// Generated by scripts/make_plcsim_bench.py. Do not edit: rerun the script.
// Recorded force-travel curves from the Python model, the evaluation recipe of the study and the
// values the NumPy evaluation gives for the same samples. Read by FB_TestBench and FB_TestPlant.
//   X, F            samples of all curves, one after the other. A curve is CurveNPull pull samples
//                   followed by the same number of return samples, in the order they were taken.
//   Case..., Exp... replay cases 1..NCases: curve, evaluation mode, expected verdict, NOK code,
//                   elements (9 per case: FpG1 FrG1 FMean FHyst FpG2 FPeak XPeak FStep XStop) and
//                   envelope counts
//   Lim             16 limits per mode, index (mode - 1) * 16 + n, n in the order
//                   G1Lo G1Hi MeanLo MeanHi HystLo HystHi RetFMin G2Lo G2Hi PeakFLo PeakFHi PeakXMin PeakXMax StepLo StopXLo StopXHi
DATA_BLOCK "DB_TestData"
{ S7_Optimized_Access := 'TRUE' }
VERSION : 0.1
NON_RETAIN
   VAR
      NCurves : Int;
      NCases : Int;
      NSamples : Int;
      Tol : Real;   // N or mm, allowed difference of an element
      GoodCurve : Int;   // curve of the good unit in the station scenario
      BadCurve : Int;   // curve of the rejected unit in the station scenario
      GateX : Real;
      Gate2X : Real;
      PeakXLo : Real;
      PeakXHi : Real;
      StepSpan : Real;
      StopF : Real;
      EnvX0 : Real;
      EnvDx : Real;
      EnvN : Int;
      CurveStart : Array[0..15] of Int;
      CurveNPull : Array[0..15] of Int;
      CaseCurve : Array[1..32] of Int;
      CaseMode : Array[1..32] of Int;
      ExpOk : Array[1..32] of Bool;
      ExpNok : Array[1..32] of Int;
      ExpEnvViol : Array[1..32] of Int;
      ExpEnvNodes : Array[1..32] of Int;
      ExpFeat : Array[0..287] of Real;
      ExpFeatValid : Array[0..287] of Bool;
      Lim : Array[0..63] of Real;
      EnvLo : Array[0..63] of Real;
      EnvHi : Array[0..63] of Real;
      X : Array[0..5931] of Real;   // mm
      F : Array[0..5931] of Real;   // N
   END_VAR

BEGIN
   NCurves := 10;
   NCases := 14;
   NSamples := 5932;
   Tol := 0.001;
   GoodCurve := 0;
   BadCurve := 6;
   GateX := 3.0;
   Gate2X := 10.0;
   PeakXLo := 13.0;
   PeakXHi := 26.0;
   StepSpan := 2.0;
   StopF := 30.0;
   EnvX0 := 1.0;
   EnvDx := 0.5;
   EnvN := 55;
   CurveStart[0] := 0;
   CurveNPull[0] := 310;
   CurveStart[1] := 620;
   CurveNPull[1] := 313;
   CurveStart[2] := 1246;
   CurveNPull[2] := 250;
   CurveStart[3] := 1746;
   CurveNPull[3] := 310;
   CurveStart[4] := 2366;
   CurveNPull[4] := 311;
   CurveStart[5] := 2988;
   CurveNPull[5] := 309;
   CurveStart[6] := 3606;
   CurveNPull[6] := 311;
   CurveStart[7] := 4228;
   CurveNPull[7] := 250;
   CurveStart[8] := 4728;
   CurveNPull[8] := 291;
   CurveStart[9] := 5310;
   CurveNPull[9] := 311;
   CaseCurve[1] := 0;
   CaseMode[1] := 3;
   ExpOk[1] := TRUE;
   ExpNok[1] := 0;
   ExpEnvViol[1] := 0;
   ExpEnvNodes[1] := 55;
   ExpFeat[0] := 6.9821014;
   ExpFeatValid[0] := TRUE;
   ExpFeat[1] := 5.37568;
   ExpFeatValid[1] := TRUE;
   ExpFeat[2] := 6.1788907;
   ExpFeatValid[2] := TRUE;
   ExpFeat[3] := 1.6064217;
   ExpFeatValid[3] := TRUE;
   ExpFeat[4] := 10.845588;
   ExpFeatValid[4] := TRUE;
   ExpFeat[5] := 16.818577;
   ExpFeatValid[5] := TRUE;
   ExpFeat[6] := 19.848608;
   ExpFeatValid[6] := TRUE;
   ExpFeat[7] := 3.9388027;
   ExpFeatValid[7] := TRUE;
   ExpFeat[8] := 29.783041;
   ExpFeatValid[8] := TRUE;
   CaseCurve[2] := 1;
   CaseMode[2] := 3;
   ExpOk[2] := TRUE;
   ExpNok[2] := 0;
   ExpEnvViol[2] := 0;
   ExpEnvNodes[2] := 55;
   ExpFeat[9] := 7.205183;
   ExpFeatValid[9] := TRUE;
   ExpFeat[10] := 5.0210447;
   ExpFeatValid[10] := TRUE;
   ExpFeat[11] := 6.113114;
   ExpFeatValid[11] := TRUE;
   ExpFeat[12] := 2.1841383;
   ExpFeatValid[12] := TRUE;
   ExpFeat[13] := 11.2528515;
   ExpFeatValid[13] := TRUE;
   ExpFeat[14] := 17.15133;
   ExpFeatValid[14] := TRUE;
   ExpFeat[15] := 18.303595;
   ExpFeatValid[15] := TRUE;
   ExpFeat[16] := 4.152199;
   ExpFeatValid[16] := TRUE;
   ExpFeat[17] := 30.096466;
   ExpFeatValid[17] := TRUE;
   CaseCurve[3] := 2;
   CaseMode[3] := 3;
   ExpNok[3] := 2;
   ExpEnvViol[3] := 43;
   ExpEnvNodes[3] := 46;
   ExpFeat[18] := 4.183258;
   ExpFeatValid[18] := TRUE;
   ExpFeat[19] := 2.565676;
   ExpFeatValid[19] := TRUE;
   ExpFeat[20] := 3.374467;
   ExpFeatValid[20] := TRUE;
   ExpFeat[21] := 1.6175817;
   ExpFeatValid[21] := TRUE;
   ExpFeat[22] := 6.124597;
   ExpFeatValid[22] := TRUE;
   ExpFeat[23] := 40.227142;
   ExpFeatValid[23] := TRUE;
   ExpFeat[24] := 23.940363;
   ExpFeatValid[24] := TRUE;
   ExpFeat[25] := 0.0;
   ExpFeatValid[25] := TRUE;
   ExpFeat[26] := 23.785864;
   ExpFeatValid[26] := TRUE;
   CaseCurve[4] := 3;
   CaseMode[4] := 3;
   ExpNok[4] := 2;
   ExpEnvViol[4] := 0;
   ExpEnvNodes[4] := 55;
   ExpFeat[27] := 5.1918726;
   ExpFeatValid[27] := TRUE;
   ExpFeat[28] := 3.556863;
   ExpFeatValid[28] := TRUE;
   ExpFeat[29] := 4.3743677;
   ExpFeatValid[29] := TRUE;
   ExpFeat[30] := 1.6350094;
   ExpFeatValid[30] := TRUE;
   ExpFeat[31] := 9.031395;
   ExpFeatValid[31] := TRUE;
   ExpFeat[32] := 14.923322;
   ExpFeatValid[32] := TRUE;
   ExpFeat[33] := 19.814;
   ExpFeatValid[33] := TRUE;
   ExpFeat[34] := 3.9026327;
   ExpFeatValid[34] := TRUE;
   ExpFeat[35] := 29.81065;
   ExpFeatValid[35] := TRUE;
   CaseCurve[5] := 4;
   CaseMode[5] := 3;
   ExpNok[5] := 2;
   ExpEnvViol[5] := 17;
   ExpEnvNodes[5] := 55;
   ExpFeat[36] := 4.6947575;
   ExpFeatValid[36] := TRUE;
   ExpFeat[37] := 3.0623243;
   ExpFeatValid[37] := TRUE;
   ExpFeat[38] := 3.8785408;
   ExpFeatValid[38] := TRUE;
   ExpFeat[39] := 1.632433;
   ExpFeatValid[39] := TRUE;
   ExpFeat[40] := 8.425375;
   ExpFeatValid[40] := TRUE;
   ExpFeat[41] := 14.073351;
   ExpFeatValid[41] := TRUE;
   ExpFeat[42] := 19.786457;
   ExpFeatValid[42] := TRUE;
   ExpFeat[43] := 3.8736982;
   ExpFeatValid[43] := TRUE;
   ExpFeat[44] := 29.815647;
   ExpFeatValid[44] := TRUE;
   CaseCurve[6] := 5;
   CaseMode[6] := 3;
   ExpNok[6] := 3;
   ExpEnvViol[6] := 41;
   ExpEnvNodes[6] := 55;
   ExpFeat[45] := 10.499536;
   ExpFeatValid[45] := TRUE;
   ExpFeat[46] := 1.8700012;
   ExpFeatValid[46] := TRUE;
   ExpFeat[47] := 6.184768;
   ExpFeatValid[47] := TRUE;
   ExpFeat[48] := 8.629534;
   ExpFeatValid[48] := TRUE;
   ExpFeat[49] := 14.390507;
   ExpFeatValid[49] := TRUE;
   ExpFeat[50] := 20.330584;
   ExpFeatValid[50] := TRUE;
   ExpFeat[51] := 19.78603;
   ExpFeatValid[51] := TRUE;
   ExpFeat[52] := 3.8881645;
   ExpFeatValid[52] := TRUE;
   ExpFeat[53] := 29.722036;
   ExpFeatValid[53] := TRUE;
   CaseCurve[7] := 6;
   CaseMode[7] := 3;
   ExpNok[7] := 5;
   ExpEnvViol[7] := 41;
   ExpEnvNodes[7] := 55;
   ExpFeat[54] := 7.0127378;
   ExpFeatValid[54] := TRUE;
   ExpFeat[55] := 5.3387175;
   ExpFeatValid[55] := TRUE;
   ExpFeat[56] := 6.175728;
   ExpFeatValid[56] := TRUE;
   ExpFeat[57] := 1.67402;
   ExpFeatValid[57] := TRUE;
   ExpFeat[58] := 7.371472;
   ExpFeatValid[58] := TRUE;
   ExpFeat[59] := 8.326099;
   ExpFeatValid[59] := TRUE;
   ExpFeat[60] := 25.861488;
   ExpFeatValid[60] := TRUE;
   ExpFeat[61] := 0.032551765;
   ExpFeatValid[61] := TRUE;
   ExpFeat[62] := 29.877676;
   ExpFeatValid[62] := TRUE;
   CaseCurve[8] := 7;
   CaseMode[8] := 3;
   ExpNok[8] := 2;
   ExpEnvViol[8] := 43;
   ExpEnvNodes[8] := 46;
   ExpFeat[63] := 4.238579;
   ExpFeatValid[63] := TRUE;
   ExpFeat[64] := 2.6031868;
   ExpFeatValid[64] := TRUE;
   ExpFeat[65] := 3.420883;
   ExpFeatValid[65] := TRUE;
   ExpFeat[66] := 1.6353921;
   ExpFeatValid[66] := TRUE;
   ExpFeat[67] := 6.187137;
   ExpFeatValid[67] := TRUE;
   ExpFeat[68] := 41.858364;
   ExpFeatValid[68] := TRUE;
   ExpFeat[69] := 23.904263;
   ExpFeatValid[69] := TRUE;
   ExpFeat[70] := 0.0;
   ExpFeatValid[70] := TRUE;
   ExpFeat[71] := 23.727392;
   ExpFeatValid[71] := TRUE;
   CaseCurve[9] := 8;
   CaseMode[9] := 3;
   ExpNok[9] := 9;
   ExpEnvViol[9] := 1;
   ExpEnvNodes[9] := 55;
   ExpFeat[72] := 7.0128746;
   ExpFeatValid[72] := TRUE;
   ExpFeat[73] := 5.3684235;
   ExpFeatValid[73] := TRUE;
   ExpFeat[74] := 6.190649;
   ExpFeatValid[74] := TRUE;
   ExpFeat[75] := 1.6444514;
   ExpFeatValid[75] := TRUE;
   ExpFeat[76] := 10.856109;
   ExpFeatValid[76] := TRUE;
   ExpFeat[77] := 16.749855;
   ExpFeatValid[77] := TRUE;
   ExpFeat[78] := 19.791138;
   ExpFeatValid[78] := TRUE;
   ExpFeat[79] := 3.8845482;
   ExpFeatValid[79] := TRUE;
   ExpFeat[80] := 27.874788;
   ExpFeatValid[80] := TRUE;
   CaseCurve[10] := 9;
   CaseMode[10] := 3;
   ExpNok[10] := 2;
   ExpEnvViol[10] := 0;
   ExpEnvNodes[10] := 55;
   ExpFeat[81] := 6.2380857;
   ExpFeatValid[81] := TRUE;
   ExpFeat[82] := 2.573432;
   ExpFeatValid[82] := TRUE;
   ExpFeat[83] := 4.405759;
   ExpFeatValid[83] := TRUE;
   ExpFeat[84] := 3.6646535;
   ExpFeatValid[84] := TRUE;
   ExpFeat[85] := 10.107543;
   ExpFeatValid[85] := TRUE;
   ExpFeat[86] := 15.954138;
   ExpFeatValid[86] := TRUE;
   ExpFeat[87] := 19.8363;
   ExpFeatValid[87] := TRUE;
   ExpFeat[88] := 3.8773146;
   ExpFeatValid[88] := TRUE;
   ExpFeat[89] := 29.792097;
   ExpFeatValid[89] := TRUE;
   CaseCurve[11] := 9;
   CaseMode[11] := 2;
   ExpOk[11] := TRUE;
   ExpNok[11] := 0;
   ExpEnvViol[11] := 0;
   ExpEnvNodes[11] := 55;
   ExpFeat[90] := 6.2380857;
   ExpFeatValid[90] := TRUE;
   ExpFeat[91] := 2.573432;
   ExpFeatValid[91] := TRUE;
   ExpFeat[92] := 4.405759;
   ExpFeatValid[92] := TRUE;
   ExpFeat[93] := 3.6646535;
   ExpFeatValid[93] := TRUE;
   ExpFeat[94] := 10.107543;
   ExpFeatValid[94] := TRUE;
   ExpFeat[95] := 15.954138;
   ExpFeatValid[95] := TRUE;
   ExpFeat[96] := 19.8363;
   ExpFeatValid[96] := TRUE;
   ExpFeat[97] := 3.8773146;
   ExpFeatValid[97] := TRUE;
   ExpFeat[98] := 29.792097;
   ExpFeatValid[98] := TRUE;
   CaseCurve[12] := 8;
   CaseMode[12] := 1;
   ExpOk[12] := TRUE;
   ExpNok[12] := 0;
   ExpEnvViol[12] := 1;
   ExpEnvNodes[12] := 55;
   ExpFeat[99] := 7.0128746;
   ExpFeatValid[99] := TRUE;
   ExpFeat[100] := 5.3684235;
   ExpFeatValid[100] := TRUE;
   ExpFeat[101] := 6.190649;
   ExpFeatValid[101] := TRUE;
   ExpFeat[102] := 1.6444514;
   ExpFeatValid[102] := TRUE;
   ExpFeat[103] := 10.856109;
   ExpFeatValid[103] := TRUE;
   ExpFeat[104] := 16.749855;
   ExpFeatValid[104] := TRUE;
   ExpFeat[105] := 19.791138;
   ExpFeatValid[105] := TRUE;
   ExpFeat[106] := 3.8845482;
   ExpFeatValid[106] := TRUE;
   ExpFeat[107] := 27.874788;
   ExpFeatValid[107] := TRUE;
   CaseCurve[13] := 0;
   CaseMode[13] := 4;
   ExpOk[13] := TRUE;
   ExpNok[13] := 0;
   ExpEnvViol[13] := 0;
   ExpEnvNodes[13] := 55;
   ExpFeat[108] := 6.9821014;
   ExpFeatValid[108] := TRUE;
   ExpFeat[109] := 5.37568;
   ExpFeatValid[109] := TRUE;
   ExpFeat[110] := 6.1788907;
   ExpFeatValid[110] := TRUE;
   ExpFeat[111] := 1.6064217;
   ExpFeatValid[111] := TRUE;
   ExpFeat[112] := 10.845588;
   ExpFeatValid[112] := TRUE;
   ExpFeat[113] := 16.818577;
   ExpFeatValid[113] := TRUE;
   ExpFeat[114] := 19.848608;
   ExpFeatValid[114] := TRUE;
   ExpFeat[115] := 3.9388027;
   ExpFeatValid[115] := TRUE;
   ExpFeat[116] := 29.783041;
   ExpFeatValid[116] := TRUE;
   CaseCurve[14] := 3;
   CaseMode[14] := 4;
   ExpOk[14] := TRUE;
   ExpNok[14] := 0;
   ExpEnvViol[14] := 0;
   ExpEnvNodes[14] := 55;
   ExpFeat[117] := 5.1918726;
   ExpFeatValid[117] := TRUE;
   ExpFeat[118] := 3.556863;
   ExpFeatValid[118] := TRUE;
   ExpFeat[119] := 4.3743677;
   ExpFeatValid[119] := TRUE;
   ExpFeat[120] := 1.6350094;
   ExpFeatValid[120] := TRUE;
   ExpFeat[121] := 9.031395;
   ExpFeatValid[121] := TRUE;
   ExpFeat[122] := 14.923322;
   ExpFeatValid[122] := TRUE;
   ExpFeat[123] := 19.814;
   ExpFeatValid[123] := TRUE;
   ExpFeat[124] := 3.9026327;
   ExpFeatValid[124] := TRUE;
   ExpFeat[125] := 29.81065;
   ExpFeatValid[125] := TRUE;
   Lim[9] := 15.241609;
   Lim[10] := 18.417305;
   Lim[16] := 5.896105;
   Lim[17] := 8.38203;
   Lim[23] := 9.4181;
   Lim[24] := 12.402887;
   Lim[25] := 14.982571;
   Lim[26] := 18.676344;
   Lim[27] := 17.139359;
   Lim[28] := 22.516165;
   Lim[29] := 2.9451215;
   Lim[30] := 28.690018;
   Lim[31] := 30.871372;
   Lim[34] := 5.186474;
   Lim[35] := 7.2080727;
   Lim[36] := -0.5455249;
   Lim[37] := 3.975223;
   Lim[38] := 1.0;
   Lim[39] := 9.212741;
   Lim[40] := 12.608247;
   Lim[41] := 14.728432;
   Lim[42] := 18.930483;
   Lim[43] := 16.769424;
   Lim[44] := 22.886099;
   Lim[45] := 2.8110514;
   Lim[46] := 28.539938;
   Lim[47] := 31.021452;
   EnvLo[0] := 4.5024867;
   EnvHi[0] := 9.917023;
   EnvLo[1] := 4.5624857;
   EnvHi[1] := 9.98225;
   EnvLo[2] := 4.530773;
   EnvHi[2] := 9.992803;
   EnvLo[3] := 4.5635424;
   EnvHi[3] := 10.004515;
   EnvLo[4] := 4.573186;
   EnvHi[4] := 10.029344;
   EnvLo[5] := 4.617667;
   EnvHi[5] := 10.026862;
   EnvLo[6] := 4.6239376;
   EnvHi[6] := 10.070514;
   EnvLo[7] := 4.670679;
   EnvHi[7] := 10.102605;
   EnvLo[8] := 4.725596;
   EnvHi[8] := 12.041139;
   EnvLo[9] := 4.700003;
   EnvHi[9] := 12.557893;
   EnvLo[10] := 4.8820324;
   EnvHi[10] := 12.779339;
   EnvLo[11] := 4.926072;
   EnvHi[11] := 12.91771;
   EnvLo[12] := 5.163019;
   EnvHi[12] := 13.360822;
   EnvLo[13] := 5.6595745;
   EnvHi[13] := 13.471234;
   EnvLo[14] := 7.878658;
   EnvHi[14] := 13.533369;
   EnvLo[15] := 8.020163;
   EnvHi[15] := 13.642666;
   EnvLo[16] := 8.08159;
   EnvHi[16] := 13.729599;
   EnvLo[17] := 8.207902;
   EnvHi[17] := 13.860825;
   EnvLo[18] := 8.30263;
   EnvHi[18] := 13.911284;
   EnvLo[19] := 8.350869;
   EnvHi[19] := 13.990431;
   EnvLo[20] := 8.425625;
   EnvHi[20] := 14.0966015;
   EnvLo[21] := 8.550419;
   EnvHi[21] := 14.182879;
   EnvLo[22] := 8.607436;
   EnvHi[22] := 14.296827;
   EnvLo[23] := 8.764787;
   EnvHi[23] := 14.390328;
   EnvLo[24] := 8.845735;
   EnvHi[24] := 14.4539795;
   EnvLo[25] := 8.9147835;
   EnvHi[25] := 14.551714;
   EnvLo[26] := 8.99205;
   EnvHi[26] := 14.698472;
   EnvLo[27] := 9.068602;
   EnvHi[27] := 15.185006;
   EnvLo[28] := 9.331687;
   EnvHi[28] := 15.688478;
   EnvLo[29] := 9.416069;
   EnvHi[29] := 16.23098;
   EnvLo[30] := 9.513143;
   EnvHi[30] := 16.795422;
   EnvLo[31] := 9.665618;
   EnvHi[31] := 17.309069;
   EnvLo[32] := 10.123489;
   EnvHi[32] := 17.854668;
   EnvLo[33] := 10.642103;
   EnvHi[33] := 18.362646;
   EnvLo[34] := 11.14989;
   EnvHi[34] := 18.931261;
   EnvLo[35] := 11.027167;
   EnvHi[35] := 18.921373;
   EnvLo[36] := 10.830289;
   EnvHi[36] := 19.396362;
   EnvLo[37] := 10.428676;
   EnvHi[37] := 19.986576;
   EnvLo[38] := 10.27112;
   EnvHi[38] := 19.496552;
   EnvLo[39] := 10.313659;
   EnvHi[39] := 19.897247;
   EnvLo[40] := 10.363278;
   EnvHi[40] := 19.346785;
   EnvLo[41] := 10.468162;
   EnvHi[41] := 18.766773;
   EnvLo[42] := 10.585302;
   EnvHi[42] := 16.553541;
   EnvLo[43] := 10.677869;
   EnvHi[43] := 16.354622;
   EnvLo[44] := 10.748317;
   EnvHi[44] := 16.457827;
   EnvLo[45] := 10.8695135;
   EnvHi[45] := 16.512941;
   EnvLo[46] := 10.998811;
   EnvHi[46] := 16.617954;
   EnvLo[47] := 11.099038;
   EnvHi[47] := 16.769545;
   EnvLo[48] := 11.214338;
   EnvHi[48] := 16.847044;
   EnvLo[49] := 11.278554;
   EnvHi[49] := 16.997396;
   EnvLo[50] := 11.41541;
   EnvHi[50] := 17.054838;
   EnvLo[51] := 11.506263;
   EnvHi[51] := 17.213253;
   EnvLo[52] := 11.623229;
   EnvHi[52] := 17.348417;
   EnvLo[53] := 11.713954;
   EnvHi[53] := 17.397055;
   EnvLo[54] := 11.844806;
   EnvHi[54] := 17.536877;
   X[1] := -0.0033742767;
   X[2] := 0.10472685;
   X[3] := 0.19745024;
   X[4] := 0.29981726;
   X[5] := 0.39700347;
   X[6] := 0.49491304;
   X[7] := 0.6008226;
   X[8] := 0.6972801;
   X[9] := 0.7991843;
   X[10] := 0.90281725;
   X[11] := 0.99573755;
   X[12] := 1.0995567;
   X[13] := 1.1978173;
   X[14] := 1.2951844;
   X[15] := 1.3980939;
   X[16] := 1.4998226;
   X[17] := 1.5985514;
   X[18] := 1.7018226;
   X[19] := 1.8003706;
   X[20] := 1.8912854;
   X[21] := 1.999562;
   X[22] := 2.0993705;
   X[23] := 2.1909237;
   X[24] := 2.2984662;
   X[25] := 2.3891046;
   X[26] := 2.4932854;
   X[27] := 2.601009;
   X[28] := 2.6959238;
   X[29] := 2.796014;
   X[30] := 2.894743;
   X[31] := 2.9955568;
   X[32] := 3.092743;
   X[33] := 3.1978333;
   X[34] := 3.292743;
   X[35] := 3.3987377;
   X[36] := 3.4987428;
   X[37] := 3.59511;
   X[38] := 3.6955674;
   X[39] := 3.7989292;
   X[40] := 3.8956633;
   X[41] := 3.9927535;
   X[42] := 4.0977483;
   X[43] := 4.197296;
   X[44] := 4.292573;
   X[45] := 4.399477;
   X[46] := 4.4931207;
   X[47] := 4.593658;
   X[48] := 4.6908493;
   X[49] := 4.7944875;
   X[50] := 4.8961205;
   X[51] := 4.9969397;
   X[52] := 5.094764;
   X[53] := 5.18994;
   X[54] := 5.2910357;
   X[55] := 5.394844;
   X[56] := 5.489573;
   X[57] := 5.5893974;
   X[58] := 5.6894984;
   X[59] := 5.7891207;
   X[60] := 5.893126;
   X[61] := 5.989312;
   X[62] := 6.076935;
   X[63] := 6.1627493;
   X[64] := 6.2443776;
   X[65] := 6.328378;
   X[66] := 6.4094586;
   X[67] := 6.5168147;
   X[68] := 6.6171765;
   X[69] := 6.718815;
   X[70] := 6.8094583;
   X[71] := 6.9220915;
   X[72] := 7.0171022;
   X[73] := 7.1126394;
   X[74] := 7.213565;
   X[75] := 7.3112035;
   X[76] := 7.4117403;
   X[77] := 7.511751;
   X[78] := 7.606661;
   X[79] := 7.708384;
   X[80] := 7.81248;
   X[81] := 7.9090276;
   X[82] := 8.005486;
   X[83] := 8.110033;
   X[84] := 8.2134;
   X[85] := 8.307496;
   X[86] := 8.410586;
   X[87] := 8.505591;
   X[88] := 8.600773;
   X[89] := 8.702959;
   X[90] := 8.809416;
   X[91] := 8.908698;
   X[92] := 8.999699;
   X[93] := 9.103602;
   X[94] := 9.201704;
   X[95] := 9.301433;
   X[96] := 9.39789;
   X[97] := 9.503613;
   X[98] := 9.601155;
   X[99] := 9.699528;
   X[100] := 9.802805;
   X[101] := 9.89989;
   X[102] := 10.003895;
   X[103] := 10.098449;
   X[104] := 10.201262;
   X[105] := 10.298172;
   X[106] := 10.399454;
   X[107] := 10.497454;
   X[108] := 10.592826;
   X[109] := 10.699917;
   X[110] := 10.798554;
   X[111] := 10.89847;
   X[112] := 10.996193;
   X[113] := 11.098837;
   X[114] := 11.192114;
   X[115] := 11.287757;
   X[116] := 11.391119;
   X[117] := 11.496119;
   X[118] := 11.592933;
   X[119] := 11.693028;
   X[120] := 11.786496;
   X[121] := 11.891943;
   X[122] := 11.991592;
   X[123] := 12.0868635;
   X[124] := 12.186582;
   X[125] := 12.291321;
   X[126] := 12.380411;
   X[127] := 12.48514;
   X[128] := 12.584327;
   X[129] := 12.683965;
   X[130] := 12.787603;
   X[131] := 12.888337;
   X[132] := 12.989885;
   X[133] := 13.08306;
   X[134] := 13.187704;
   X[135] := 13.284523;
   X[136] := 13.3848;
   X[137] := 13.487896;
   X[138] := 13.587353;
   X[139] := 13.678811;
   X[140] := 13.784454;
   X[141] := 13.882715;
   X[142] := 13.981008;
   X[143] := 14.078545;
   X[144] := 14.183087;
   X[145] := 14.28164;
   X[146] := 14.38038;
   X[147] := 14.475013;
   X[148] := 14.574927;
   X[149] := 14.682922;
   X[150] := 14.780104;
   X[151] := 14.878199;
   X[152] := 14.975023;
   X[153] := 15.076039;
   X[154] := 15.17287;
   X[155] := 15.271434;
   X[156] := 15.363907;
   X[157] := 15.460098;
   X[158] := 15.557104;
   X[159] := 15.660487;
   X[160] := 15.751045;
   X[161] := 15.851062;
   X[162] := 15.951705;
   X[163] := 16.053541;
   X[164] := 16.149647;
   X[165] := 16.244019;
   X[166] := 16.34385;
   X[167] := 16.440685;
   X[168] := 16.537062;
   X[169] := 16.62862;
   X[170] := 16.734083;
   X[171] := 16.83637;
   X[172] := 16.92229;
   X[173] := 17.019585;
   X[174] := 17.119505;
   X[175] := 17.217972;
   X[176] := 17.316803;
   X[177] := 17.418;
   X[178] := 17.508282;
   X[179] := 17.611292;
   X[180] := 17.70858;
   X[181] := 17.800692;
   X[182] := 17.902872;
   X[183] := 17.99408;
   X[184] := 18.09909;
   X[185] := 18.191565;
   X[186] := 18.287483;
   X[187] := 18.387772;
   X[188] := 18.49033;
   X[189] := 18.585798;
   X[190] := 18.676447;
   X[191] := 18.777182;
   X[192] := 18.874111;
   X[193] := 18.979118;
   X[194] := 19.070032;
   X[195] := 19.165964;
   X[196] := 19.270985;
   X[197] := 19.360996;
   X[198] := 19.462011;
   X[199] := 19.55457;
   X[200] := 19.65848;
   X[201] := 19.755777;
   X[202] := 19.848608;
   X[203] := 19.970793;
   X[204] := 20.087416;
   X[205] := 20.211292;
   X[206] := 20.32783;
   X[207] := 20.445093;
   X[208] := 20.557806;
   X[209] := 20.648077;
   X[210] := 20.741636;
   X[211] := 20.84809;
   X[212] := 20.953089;
   X[213] := 21.043913;
   X[214] := 21.147093;
   X[215] := 21.24119;
   X[216] := 21.348913;
   X[217] := 21.449648;
   X[218] := 21.545195;
   X[219] := 21.634748;
   X[220] := 21.745749;
   X[221] := 21.841301;
   X[222] := 21.946121;
   X[223] := 22.040205;
   X[224] := 22.143402;
   X[225] := 22.240217;
   X[226] := 22.341042;
   X[227] := 22.44068;
   X[228] := 22.53859;
   X[229] := 22.634499;
   X[230] := 22.738136;
   X[231] := 22.838509;
   X[232] := 22.941322;
   X[233] := 23.042967;
   X[234] := 23.129976;
   X[235] := 23.239418;
   X[236] := 23.335434;
   X[237] := 23.430067;
   X[238] := 23.531801;
   X[239] := 23.641802;
   X[240] := 23.734535;
   X[241] := 23.835356;
   X[242] := 23.933903;
   X[243] := 24.02927;
   X[244] := 24.133179;
   X[245] := 24.232546;
   X[246] := 24.332918;
   X[247] := 24.43128;
   X[248] := 24.52801;
   X[249] := 24.624918;
   X[250] := 24.728653;
   X[251] := 24.823557;
   X[252] := 24.925116;
   X[253] := 25.026297;
   X[254] := 25.123116;
   X[255] := 25.230398;
   X[256] := 25.325674;
   X[257] := 25.426765;
   X[258] := 25.523584;
   X[259] := 25.621408;
   X[260] := 25.71895;
   X[261] := 25.820227;
   X[262] := 25.919882;
   X[263] := 26.019594;
   X[264] := 26.116701;
   X[265] := 26.216702;
   X[266] := 26.315063;
   X[267] := 26.42161;
   X[268] := 26.524881;
   X[269] := 26.622345;
   X[270] := 26.714718;
   X[271] := 26.815802;
   X[272] := 26.917803;
   X[273] := 27.014627;
   X[274] := 27.115812;
   X[275] := 27.214813;
   X[276] := 27.312366;
   X[277] := 27.413908;
   X[278] := 27.51119;
   X[279] := 27.612286;
   X[280] := 27.709558;
   X[281] := 27.811739;
   X[282] := 27.911112;
   X[283] := 28.007027;
   X[284] := 28.111387;
   X[285] := 28.199669;
   X[286] := 28.301207;
   X[287] := 28.40676;
   X[288] := 28.508398;
   X[289] := 28.60403;
   X[290] := 28.701595;
   X[291] := 28.8095;
   X[292] := 28.900776;
   X[293] := 29.00051;
   X[294] := 29.101877;
   X[295] := 29.200064;
   X[296] := 29.301426;
   X[297] := 29.398798;
   X[298] := 29.500973;
   X[299] := 29.572319;
   X[300] := 29.6092;
   X[301] := 29.646812;
   X[302] := 29.686869;
   X[303] := 29.716297;
   X[304] := 29.758177;
   X[305] := 29.799242;
   X[306] := 29.837845;
   X[307] := 29.867996;
   X[308] := 29.91243;
   X[309] := 29.94758;
   X[310] := 29.943314;
   X[311] := 29.928886;
   X[312] := 29.886644;
   X[313] := 29.850302;
   X[314] := 29.813248;
   X[315] := 29.77291;
   X[316] := 29.739481;
   X[317] := 29.693878;
   X[318] := 29.666807;
   X[319] := 29.625662;
   X[320] := 29.588596;
   X[321] := 29.545658;
   X[322] := 29.446291;
   X[323] := 29.346828;
   X[324] := 29.248291;
   X[325] := 29.144827;
   X[326] := 29.049004;
   X[327] := 28.937727;
   X[328] := 28.847637;
   X[329] := 28.75453;
   X[330] := 28.642721;
   X[331] := 28.549807;
   X[332] := 28.448168;
   X[333] := 28.348167;
   X[334] := 28.251705;
   X[335] := 28.151072;
   X[336] := 28.05543;
   X[337] := 27.9487;
   X[338] := 27.857418;
   X[339] := 27.751062;
   X[340] := 27.654417;
   X[341] := 27.556412;
   X[342] := 27.45969;
   X[343] := 27.360954;
   X[344] := 27.257498;
   X[345] := 27.15513;
   X[346] := 27.059216;
   X[347] := 26.958311;
   X[348] := 26.85785;
   X[349] := 26.761482;
   X[350] := 26.654758;
   X[351] := 26.5573;
   X[352] := 26.460743;
   X[353] := 26.360561;
   X[354] := 26.257103;
   X[355] := 26.160013;
   X[356] := 26.06664;
   X[357] := 25.96328;
   X[358] := 25.863731;
   X[359] := 25.76454;
   X[360] := 25.668083;
   X[361] := 25.56563;
   X[362] := 25.464897;
   X[363] := 25.367987;
   X[364] := 25.26344;
   X[365] := 25.167982;
   X[366] := 25.070257;
   X[367] := 24.966524;
   X[368] := 24.871796;
   X[369] := 24.767876;
   X[370] := 24.67279;
   X[371] := 24.576056;
   X[372] := 24.471146;
   X[373] := 24.368502;
   X[374] := 24.26669;
   X[375] := 24.170046;
   X[376] := 24.073677;
   X[377] := 23.97786;
   X[378] := 23.87113;
   X[379] := 23.777668;
   X[380] := 23.676853;
   X[381] := 23.576395;
   X[382] := 23.480204;
   X[383] := 23.375023;
   X[384] := 23.272934;
   X[385] := 23.17702;
   X[386] := 23.081102;
   X[387] := 22.978556;
   X[388] := 22.88028;
   X[389] := 22.779646;
   X[390] := 22.677635;
   X[391] := 22.582449;
   X[392] := 22.482183;
   X[393] := 22.376087;
   X[394] := 22.28681;
   X[395] := 22.185173;
   X[396] := 22.084444;
   X[397] := 21.981167;
   X[398] := 21.891161;
   X[399] := 21.780619;
   X[400] := 21.684343;
   X[401] := 21.589523;
   X[402] := 21.48388;
   X[403] := 21.391508;
   X[404] := 21.285975;
   X[405] := 21.187326;
   X[406] := 21.08787;
   X[407] := 20.986044;
   X[408] := 20.88931;
   X[409] := 20.790411;
   X[410] := 20.692492;
   X[411] := 20.591034;
   X[412] := 20.4904;
   X[413] := 20.394842;
   X[414] := 20.293018;
   X[415] := 20.197294;
   X[416] := 20.102022;
   X[417] := 19.994108;
   X[418] := 19.893831;
   X[419] := 19.797018;
   X[420] := 19.694916;
   X[421] := 19.590475;
   X[422] := 19.501102;
   X[423] := 19.397188;
   X[424] := 19.298725;
   X[425] := 19.19691;
   X[426] := 19.100178;
   X[427] := 18.99881;
   X[428] := 18.902714;
   X[429] := 18.797997;
   X[430] := 18.700708;
   X[431] := 18.604261;
   X[432] := 18.502884;
   X[433] := 18.39889;
   X[434] := 18.303162;
   X[435] := 18.206156;
   X[436] := 18.103241;
   X[437] := 17.99897;
   X[438] := 17.907688;
   X[439] := 17.802235;
   X[440] := 17.704773;
   X[441] := 17.608416;
   X[442] := 17.508411;
   X[443] := 17.407219;
   X[444] := 17.30849;
   X[445] := 17.209394;
   X[446] := 17.109943;
   X[447] := 17.011847;
   X[448] := 16.906948;
   X[449] := 16.809395;
   X[450] := 16.708118;
   X[451] := 16.613565;
   X[452] := 16.507107;
   X[453] := 16.412107;
   X[454] := 16.31701;
   X[455] := 16.208832;
   X[456] := 16.112278;
   X[457] := 16.011374;
   X[458] := 15.918001;
   X[459] := 15.814639;
   X[460] := 15.7179;
   X[461] := 15.617182;
   X[462] := 15.515448;
   X[463] := 15.413996;
   X[464] := 15.3189;
   X[465] := 15.21989;
   X[466] := 15.117075;
   X[467] := 15.018708;
   X[468] := 14.91516;
   X[469] := 14.81798;
   X[470] := 14.721788;
   X[471] := 14.619889;
   X[472] := 14.519878;
   X[473] := 14.4160595;
   X[474] := 14.324873;
   X[475] := 14.220602;
   X[476] := 14.128693;
   X[477] := 14.019857;
   X[478] := 13.914687;
   X[479] := 13.827314;
   X[480] := 13.7215;
   X[481] := 13.626677;
   X[482] := 13.521501;
   X[483] := 13.424581;
   X[484] := 13.327847;
   X[485] := 13.228756;
   X[486] := 13.133394;
   X[487] := 13.029112;
   X[488] := 12.930293;
   X[489] := 12.828841;
   X[490] := 12.727287;
   X[491] := 12.62883;
   X[492] := 12.531464;
   X[493] := 12.429921;
   X[494] := 12.327181;
   X[495] := 12.229639;
   X[496] := 12.131453;
   X[497] := 12.032723;
   X[498] := 11.925458;
   X[499] := 11.833815;
   X[500] := 11.732442;
   X[501] := 11.633894;
   X[502] := 11.536803;
   X[503] := 11.433075;
   X[504] := 11.328346;
   X[505] := 11.23716;
   X[506] := 11.135245;
   X[507] := 11.032245;
   X[508] := 10.939425;
   X[509] := 10.837878;
   X[510] := 10.737963;
   X[511] := 10.632873;
   X[512] := 10.537234;
   X[513] := 10.437139;
   X[514] := 10.339868;
   X[515] := 10.24041;
   X[516] := 10.143681;
   X[517] := 10.045037;
   X[518] := 9.939037;
   X[519] := 9.833128;
   X[520] := 9.744676;
   X[521] := 9.642303;
   X[522] := 9.540303;
   X[523] := 9.441941;
   X[524] := 9.343032;
   X[525] := 9.2415695;
   X[526] := 9.141931;
   X[527] := 9.047192;
   X[528] := 8.943649;
   X[529] := 8.843558;
   X[530] := 8.747462;
   X[531] := 8.645282;
   X[532] := 8.554914;
   X[533] := 8.446638;
   X[534] := 8.344186;
   X[535] := 8.247452;
   X[536] := 8.145633;
   X[537] := 8.051356;
   X[538] := 7.9505424;
   X[539] := 7.854803;
   X[540] := 7.749255;
   X[541] := 7.6534357;
   X[542] := 7.5542603;
   X[543] := 7.453893;
   X[544] := 7.3493347;
   X[545] := 7.2504253;
   X[546] := 7.1519732;
   X[547] := 7.054606;
   X[548] := 6.9581485;
   X[549] := 6.8538775;
   X[550] := 6.7531433;
   X[551] := 6.657409;
   X[552] := 6.5563293;
   X[553] := 6.4607816;
   X[554] := 6.3632812;
   X[555] := 6.274286;
   X[556] := 6.1935673;
   X[557] := 6.108753;
   X[558] := 6.03021;
   X[559] := 5.9339066;
   X[560] := 5.8310876;
   X[561] := 5.731545;
   X[562] := 5.6369066;
   X[563] := 5.531364;
   X[564] := 5.437353;
   X[565] := 5.337811;
   X[566] := 5.2275395;
   X[567] := 5.126901;
   X[568] := 5.03872;
   X[569] := 4.9384384;
   X[570] := 4.8375287;
   X[571] := 4.739082;
   X[572] := 4.634901;
   X[573] := 4.5331616;
   X[574] := 4.4404383;
   X[575] := 4.329167;
   X[576] := 4.233348;
   X[577] := 4.1344438;
   X[578] := 4.0365286;
   X[579] := 3.9392576;
   X[580] := 3.834167;
   X[581] := 3.7369862;
   X[582] := 3.633433;
   X[583] := 3.5345287;
   X[584] := 3.4394383;
   X[585] := 3.3372576;
   X[586] := 3.2332575;
   X[587] := 3.140433;
   X[588] := 3.043066;
   X[589] := 2.9320712;
   X[590] := 2.8413372;
   X[591] := 2.7396085;
   X[592] := 2.6366086;
   X[593] := 2.5347893;
   X[594] := 2.441518;
   X[595] := 2.342518;
   X[596] := 2.2378001;
   X[597] := 2.1382415;
   X[598] := 2.034066;
   X[599] := 1.9376031;
   X[600] := 1.8358798;
   X[601] := 1.7395127;
   X[602] := 1.6385127;
   X[603] := 1.540151;
   X[604] := 1.4401511;
   X[605] := 1.3368851;
   X[606] := 1.2400553;
   X[607] := 1.133151;
   X[608] := 1.0449648;
   X[609] := 0.939784;
   X[610] := 0.8416882;
   X[611] := 0.7337893;
   X[612] := 0.6410499;
   X[613] := 0.5402415;
   X[614] := 0.43896484;
   X[615] := 0.34032118;
   X[616] := 0.23696484;
   X[617] := 0.14223076;
   X[618] := 0.03723076;
   X[619] := 0.07943374;
   X[621] := 0.058969617;
   X[622] := 0.1601451;
   X[623] := 0.25842172;
   X[624] := 0.36087385;
   X[625] := 0.45877805;
   X[626] := 0.5548792;
   X[627] := 0.6574271;
   X[628] := 0.75815046;
   X[629] := 0.85487384;
   X[630] := 0.9517888;
   X[631] := 1.053975;
   X[632] := 1.1582409;
   X[633] := 1.2541559;
   X[634] := 1.3572463;
   X[635] := 1.4556025;
   X[636] := 1.5523367;
   X[637] := 1.6556187;
   X[638] := 1.7556983;
   X[639] := 1.8526186;
   X[640] := 1.9547037;
   X[641] := 2.0571558;
   X[642] := 2.1517036;
   X[643] := 2.2567995;
   X[644] := 2.3577092;
   X[645] := 2.4552517;
   X[646] := 2.5556185;
   X[647] := 2.6554377;
   X[648] := 2.7547994;
   X[649] := 2.850161;
   X[650] := 2.9497144;
   X[651] := 3.0517995;
   X[652] := 3.1496186;
   X[653] := 3.257076;
   X[654] := 3.3558953;
   X[655] := 3.4521666;
   X[656] := 3.5518048;
   X[657] := 3.653624;
   X[658] := 3.7534378;
   X[659] := 3.852991;
   X[660] := 3.9552622;
   X[661] := 4.04972;
   X[662] := 4.1526294;
   X[663] := 4.255996;
   X[664] := 4.3528047;
   X[665] := 4.4510016;
   X[666] := 4.5480866;
   X[667] := 4.6492677;
   X[668] := 4.7482677;
   X[669] := 4.853805;
   X[670] := 4.9477253;
   X[671] := 5.051906;
   X[672] := 5.151358;
   X[673] := 5.2348957;
   X[674] := 5.3198113;
   X[675] := 5.4007053;
   X[676] := 5.4895253;
   X[677] := 5.573419;
   X[678] := 5.673228;
   X[679] := 5.771866;
   X[680] := 5.871143;
   X[681] := 5.969329;
   X[682] := 6.072978;
   X[683] := 6.165616;
   X[684] := 6.2763395;
   X[685] := 6.37834;
   X[686] := 6.4693394;
   X[687] := 6.5714407;
   X[688] := 6.6652493;
   X[689] := 6.770627;
   X[690] := 6.8630843;
   X[691] := 6.9633555;
   X[692] := 7.0697227;
   X[693] := 7.168909;
   X[694] := 7.2685523;
   X[695] := 7.3637385;
   X[696] := 7.4669037;
   X[697] := 7.563648;
   X[698] := 7.6645527;
   X[699] := 7.7610154;
   X[700] := 7.8674674;
   X[701] := 7.9631057;
   X[702] := 8.063478;
   X[703] := 8.159749;
   X[704] := 8.254574;
   X[705] := 8.355664;
   X[706] := 8.462856;
   X[707] := 8.553574;
   X[708] := 8.662393;
   X[709] := 8.762766;
   X[710] := 8.8588505;
   X[711] := 8.952951;
   X[712] := 9.056047;
   X[713] := 9.15259;
   X[714] := 9.251148;
   X[715] := 9.357691;
   X[716] := 9.453968;
   X[717] := 9.555329;
   X[718] := 9.654702;
   X[719] := 9.75134;
   X[720] := 9.855978;
   X[721] := 9.954888;
   X[722] := 10.04817;
   X[723] := 10.15099;
   X[724] := 10.252255;
   X[725] := 10.3547125;
   X[726] := 10.451904;
   X[727] := 10.551271;
   X[728] := 10.646809;
   X[729] := 10.748909;
   X[730] := 10.853186;
   X[731] := 10.952457;
   X[732] := 11.050553;
   X[733] := 11.14801;
   X[734] := 11.246378;
   X[735] := 11.350468;
   X[736] := 11.444835;
   X[737] := 11.546383;
   X[738] := 11.644745;
   X[739] := 11.748659;
   X[740] := 11.844665;
   X[741] := 11.942393;
   X[742] := 12.038213;
   X[743] := 12.13958;
   X[744] := 12.245122;
   X[745] := 12.339048;
   X[746] := 12.439409;
   X[747] := 12.540957;
   X[748] := 12.639862;
   X[749] := 12.740053;
   X[750] := 12.837516;
   X[751] := 12.932607;
   X[752] := 13.040059;
   X[753] := 13.139059;
   X[754] := 13.238154;
   X[755] := 13.338431;
   X[756] := 13.4359;
   X[757] := 13.5304575;
   X[758] := 13.635559;
   X[759] := 13.72675;
   X[760] := 13.818857;
   X[761] := 13.918681;
   X[762] := 14.016246;
   X[763] := 14.117352;
   X[764] := 14.217459;
   X[765] := 14.311023;
   X[766] := 14.407762;
   X[767] := 14.50431;
   X[768] := 14.610332;
   X[769] := 14.701975;
   X[770] := 14.796544;
   X[771] := 14.899007;
   X[772] := 14.994475;
   X[773] := 15.085858;
   X[774] := 15.194316;
   X[775] := 15.28988;
   X[776] := 15.3827095;
   X[777] := 15.478273;
   X[778] := 15.579289;
   X[779] := 15.676763;
   X[780] := 15.776773;
   X[781] := 15.875156;
   X[782] := 15.973704;
   X[783] := 16.068811;
   X[784] := 16.163736;
   X[785] := 16.2553;
   X[786] := 16.359764;
   X[787] := 16.457323;
   X[788] := 16.552242;
   X[789] := 16.653168;
   X[790] := 16.743004;
   X[791] := 16.841015;
   X[792] := 16.939758;
   X[793] := 17.037136;
   X[794] := 17.140327;
   X[795] := 17.235802;
   X[796] := 17.331541;
   X[797] := 17.428104;
   X[798] := 17.52593;
   X[799] := 17.631126;
   X[800] := 17.718876;
   X[801] := 17.81943;
   X[802] := 17.915802;
   X[803] := 18.00819;
   X[804] := 18.111834;
   X[805] := 18.202488;
   X[806] := 18.303595;
   X[807] := 18.407286;
   X[808] := 18.52944;
   X[809] := 18.65905;
   X[810] := 18.7763;
   X[811] := 18.901001;
   X[812] := 19.0094;
   X[813] := 19.106045;
   X[814] := 19.20614;
   X[815] := 19.303415;
   X[816] := 19.40779;
   X[817] := 19.507235;
   X[818] := 19.609697;
   X[819] := 19.70224;
   X[820] := 19.802341;
   X[821] := 19.900156;
   X[822] := 20.002895;
   X[823] := 20.102533;
   X[824] := 20.202618;
   X[825] := 20.304895;
   X[826] := 20.402363;
   X[827] := 20.497267;
   X[828] := 20.599997;
   X[829] := 20.69355;
   X[830] := 20.796188;
   X[831] := 20.893097;
   X[832] := 20.992193;
   X[833] := 21.097012;
   X[834] := 21.191204;
   X[835] := 21.29547;
   X[836] := 21.400927;
   X[837] := 21.492119;
   X[838] := 21.598661;
   X[839] := 21.689854;
   X[840] := 21.794113;
   X[841] := 21.885592;
   X[842] := 21.988316;
   X[843] := 22.08878;
   X[844] := 22.190773;
   X[845] := 22.293049;
   X[846] := 22.38805;
   X[847] := 22.484604;
   X[848] := 22.585506;
   X[849] := 22.687784;
   X[850] := 22.784433;
   X[851] := 22.885614;
   X[852] := 22.98833;
   X[853] := 23.082354;
   X[854] := 23.185162;
   X[855] := 23.283348;
   X[856] := 23.381716;
   X[857] := 23.482725;
   X[858] := 23.583992;
   X[859] := 23.68372;
   X[860] := 23.78337;
   X[861] := 23.879997;
   X[862] := 23.972647;
   X[863] := 24.07764;
   X[864] := 24.179012;
   X[865] := 24.279741;
   X[866] := 24.376842;
   X[867] := 24.48021;
   X[868] := 24.577572;
   X[869] := 24.6793;
   X[870] := 24.773943;
   X[871] := 24.874945;
   X[872] := 24.974407;
   X[873] := 25.07404;
   X[874] := 25.175955;
   X[875] := 25.274588;
   X[876] := 25.366964;
   X[877] := 25.468056;
   X[878] := 25.566055;
   X[879] := 25.66897;
   X[880] := 25.770609;
   X[881] := 25.869247;
   X[882] := 25.965885;
   X[883] := 26.0708;
   X[884] := 26.170258;
   X[885] := 26.2708;
   X[886] := 26.36344;
   X[887] := 26.460264;
   X[888] := 26.56645;
   X[889] := 26.666822;
   X[890] := 26.763725;
   X[891] := 26.867178;
   X[892] := 26.958647;
   X[893] := 27.05411;
   X[894] := 27.163929;
   X[895] := 27.263475;
   X[896] := 27.364023;
   X[897] := 27.460024;
   X[898] := 27.559578;
   X[899] := 27.659397;
   X[900] := 27.761215;
   X[901] := 27.85913;
   X[902] := 27.956684;
   X[903] := 28.054413;
   X[904] := 28.157417;
   X[905] := 28.249779;
   X[906] := 28.357328;
   X[907] := 28.453423;
   X[908] := 28.551237;
   X[909] := 28.653881;
   X[910] := 28.746983;
   X[911] := 28.850885;
   X[912] := 28.955158;
   X[913] := 29.047626;
   X[914] := 29.149813;
   X[915] := 29.249632;
   X[916] := 29.350636;
   X[917] := 29.44836;
   X[918] := 29.546822;
   X[919] := 29.64455;
   X[920] := 29.74519;
   X[921] := 29.845291;
   X[922] := 29.898531;
   X[923] := 29.932146;
   X[924] := 29.975742;
   X[925] := 30.014538;
   X[926] := 30.052784;
   X[927] := 30.09384;
   X[928] := 30.124363;
   X[929] := 30.161966;
   X[930] := 30.199852;
   X[931] := 30.23428;
   X[932] := 30.276073;
   X[933] := 30.279707;
   X[934] := 30.259258;
   X[935] := 30.220552;
   X[936] := 30.182497;
   X[937] := 30.147161;
   X[938] := 30.109282;
   X[939] := 30.07712;
   X[940] := 30.027245;
   X[941] := 29.995913;
   X[942] := 29.958479;
   X[943] := 29.921057;
   X[944] := 29.88163;
   X[945] := 29.803432;
   X[946] := 29.702337;
   X[947] := 29.604788;
   X[948] := 29.508512;
   X[949] := 29.404512;
   X[950] := 29.309692;
   X[951] := 29.208055;
   X[952] := 29.105412;
   X[953] := 29.010315;
   X[954] := 28.907495;
   X[955] := 28.810219;
   X[956] := 28.708496;
   X[957] := 28.606033;
   X[958] := 28.511213;
   X[959] := 28.409018;
   X[960] := 28.308836;
   X[961] := 28.206108;
   X[962] := 28.11083;
   X[963] := 28.009554;
   X[964] := 27.920464;
   X[965] := 27.817097;
   X[966] := 27.714096;
   X[967] := 27.614098;
   X[968] := 27.519081;
   X[969] := 27.421623;
   X[970] := 27.311539;
   X[971] := 27.215809;
   X[972] := 27.113165;
   X[973] := 27.011442;
   X[974] := 26.923613;
   X[975] := 26.819523;
   X[976] := 26.72316;
   X[977] := 26.624512;
   X[978] := 26.518154;
   X[979] := 26.424501;
   X[980] := 26.324501;
   X[981] := 26.223682;
   X[982] := 26.12832;
   X[983] := 26.023682;
   X[984] := 25.925581;
   X[985] := 25.826756;
   X[986] := 25.725304;
   X[987] := 25.633213;
   X[988] := 25.526209;
   X[989] := 25.431484;
   X[990] := 25.327932;
   X[991] := 25.231379;
   X[992] := 25.124107;
   X[993] := 25.027378;
   X[994] := 24.92774;
   X[995] := 24.827005;
   X[996] := 24.72682;
   X[997] := 24.634266;
   X[998] := 24.533634;
   X[999] := 24.435629;
   X[1000] := 24.333357;
   X[1001] := 24.235714;
   X[1002] := 24.134075;
   X[1003] := 24.037159;
   X[1004] := 23.934883;
   X[1005] := 23.83689;
   X[1006] := 23.733522;
   X[1007] := 23.644058;
   X[1008] := 23.538336;
   X[1009] := 23.439335;
   X[1010] := 23.337143;
   X[1011] := 23.241873;
   X[1012] := 23.141325;
   X[1013] := 23.039495;
   X[1014] := 22.943308;
   X[1015] := 22.836676;
   X[1016] := 22.740585;
   X[1017] := 22.643122;
   X[1018] := 22.548845;
   X[1019] := 22.443756;
   X[1020] := 22.34893;
   X[1021] := 22.245022;
   X[1022] := 22.14148;
   X[1023] := 22.045925;
   X[1024] := 21.948095;
   X[1025] := 21.845825;
   X[1026] := 21.747463;
   X[1027] := 21.648638;
   X[1028] := 21.544724;
   X[1029] := 21.452633;
   X[1030] := 21.34591;
   X[1031] := 21.252352;
   X[1032] := 21.149809;
   X[1033] := 21.053707;
   X[1034] := 20.957075;
   X[1035] := 20.850708;
   X[1036] := 20.75434;
   X[1037] := 20.64933;
   X[1038] := 20.556244;
   X[1039] := 20.450605;
   X[1040] := 20.35551;
   X[1041] := 20.255686;
   X[1042] := 20.158957;
   X[1043] := 20.061596;
   X[1044] := 19.960772;
   X[1045] := 19.857952;
   X[1046] := 19.762127;
   X[1047] := 19.659489;
   X[1048] := 19.561398;
   X[1049] := 19.463669;
   X[1050] := 19.359297;
   X[1051] := 19.259573;
   X[1052] := 19.161749;
   X[1053] := 19.060844;
   X[1054] := 18.962467;
   X[1055] := 18.862371;
   X[1056] := 18.765282;
   X[1057] := 18.660913;
   X[1058] := 18.566366;
   X[1059] := 18.460653;
   X[1060] := 18.360914;
   X[1061] := 18.270807;
   X[1062] := 18.172451;
   X[1063] := 18.065079;
   X[1064] := 17.969627;
   X[1065] := 17.871622;
   X[1066] := 17.768164;
   X[1067] := 17.67243;
   X[1068] := 17.567436;
   X[1069] := 17.47643;
   X[1070] := 17.368792;
   X[1071] := 17.271786;
   X[1072] := 17.17751;
   X[1073] := 17.071148;
   X[1074] := 16.969872;
   X[1075] := 16.872866;
   X[1076] := 16.770239;
   X[1077] := 16.681765;
   X[1078] := 16.574047;
   X[1079] := 16.477217;
   X[1080] := 16.370668;
   X[1081] := 16.275764;
   X[1082] := 16.177212;
   X[1083] := 16.073658;
   X[1084] := 15.979759;
   X[1085] := 15.87902;
   X[1086] := 15.777563;
   X[1087] := 15.671382;
   X[1088] := 15.586376;
   X[1089] := 15.481924;
   X[1090] := 15.379919;
   X[1091] := 15.276377;
   X[1092] := 15.181281;
   X[1093] := 15.08636;
   X[1094] := 14.982185;
   X[1095] := 14.887541;
   X[1096] := 14.778909;
   X[1097] := 14.685083;
   X[1098] := 14.590627;
   X[1099] := 14.482345;
   X[1100] := 14.385892;
   X[1101] := 14.288073;
   X[1102] := 14.186977;
   X[1103] := 14.087796;
   X[1104] := 13.983977;
   X[1105] := 13.882429;
   X[1106] := 13.788419;
   X[1107] := 13.691237;
   X[1108] := 13.585786;
   X[1109] := 13.489599;
   X[1110] := 13.390775;
   X[1111] := 13.289956;
   X[1112] := 13.196493;
   X[1113] := 13.09286;
   X[1114] := 12.993312;
   X[1115] := 12.887945;
   X[1116] := 12.791126;
   X[1117] := 12.695663;
   X[1118] := 12.598573;
   X[1119] := 12.4952965;
   X[1120] := 12.398929;
   X[1121] := 12.295924;
   X[1122] := 12.19511;
   X[1123] := 12.095748;
   X[1124] := 11.997562;
   X[1125] := 11.899285;
   X[1126] := 11.795099;
   X[1127] := 11.700924;
   X[1128] := 11.59928;
   X[1129] := 11.501275;
   X[1130] := 11.400998;
   X[1131] := 11.296269;
   X[1132] := 11.20136;
   X[1133] := 11.098631;
   X[1134] := 10.997439;
   X[1135] := 10.901258;
   X[1136] := 10.802343;
   X[1137] := 10.704705;
   X[1138] := 10.604073;
   X[1139] := 10.503344;
   X[1140] := 10.405062;
   X[1141] := 10.304508;
   X[1142] := 10.20687;
   X[1143] := 10.110237;
   X[1144] := 10.015503;
   X[1145] := 9.908232;
   X[1146] := 9.80387;
   X[1147] := 9.70986;
   X[1148] := 9.613317;
   X[1149] := 9.510488;
   X[1150] := 9.412759;
   X[1151] := 9.315125;
   X[1152] := 9.2118435;
   X[1153] := 9.115025;
   X[1154] := 9.007386;
   X[1155] := 8.917743;
   X[1156] := 8.812657;
   X[1157] := 8.711567;
   X[1158] := 8.614014;
   X[1159] := 8.5132;
   X[1160] := 8.413094;
   X[1161] := 8.316461;
   X[1162] := 8.2181835;
   X[1163] := 8.115466;
   X[1164] := 8.0167265;
   X[1165] := 7.91754;
   X[1166] := 7.821811;
   X[1167] := 7.720806;
   X[1168] := 7.614529;
   X[1169] := 7.5185294;
   X[1170] := 7.415439;
   X[1171] := 7.320343;
   X[1172] := 7.2262526;
   X[1173] := 7.1214337;
   X[1174] := 7.015976;
   X[1175] := 6.92479;
   X[1176] := 6.824875;
   X[1177] := 6.7247844;
   X[1178] := 6.624508;
   X[1179] := 6.5194283;
   X[1180] := 6.4205985;
   X[1181] := 6.325327;
   X[1182] := 6.2258644;
   X[1183] := 6.1244917;
   X[1184] := 6.02304;
   X[1185] := 5.9274974;
   X[1186] := 5.825758;
   X[1187] := 5.7219496;
   X[1188] := 5.6314015;
   X[1189] := 5.536194;
   X[1190] := 5.44547;
   X[1191] := 5.3669214;
   X[1192] := 5.285751;
   X[1193] := 5.202383;
   X[1194] := 5.105436;
   X[1195] := 5.006702;
   X[1196] := 4.9036064;
   X[1197] := 4.806521;
   X[1198] := 4.706877;
   X[1199] := 4.6049786;
   X[1200] := 4.5074253;
   X[1201] := 4.4004254;
   X[1202] := 4.30834;
   X[1203] := 4.207973;
   X[1204] := 4.1086006;
   X[1205] := 4.004883;
   X[1206] := 3.9012392;
   X[1207] := 3.8079624;
   X[1208] := 3.7125103;
   X[1209] := 3.6096008;
   X[1210] := 3.5041487;
   X[1211] := 3.413053;
   X[1212] := 3.30342;
   X[1213] := 3.21142;
   X[1214] := 3.1053243;
   X[1215] := 3.0126913;
   X[1216] := 2.9129572;
   X[1217] := 2.8093243;
   X[1218] := 2.699053;
   X[1219] := 2.6135051;
   X[1220] := 2.506138;
   X[1221] := 2.4069571;
   X[1222] := 2.3082337;
   X[1223] := 2.2100475;
   X[1224] := 2.1109626;
   X[1225] := 2.00642;
   X[1226] := 1.910505;
   X[1227] := 1.8110476;
   X[1228] := 1.7060529;
   X[1229] := 1.6115955;
   X[1230] := 1.5136752;
   X[1231] := 1.4113135;
   X[1232] := 1.3050423;
   X[1233] := 1.2158561;
   X[1234] := 1.1087602;
   X[1235] := 1.0117602;
   X[1236] := 0.9073135;
   X[1237] := 0.8141273;
   X[1238] := 0.7076752;
   X[1239] := 0.6063986;
   X[1240] := 0.50649434;
   X[1241] := 0.40968055;
   X[1242] := 0.31476563;
   X[1243] := 0.20966984;
   X[1244] := 0.11121774;
   X[1245] := 0.008217737;
   X[1247] := 0.08626114;
   X[1248] := 0.16408622;
   X[1249] := 0.25262398;
   X[1250] := 0.34693274;
   X[1251] := 0.44683695;
   X[1252] := 0.5450178;
   X[1253] := 0.64548063;
   X[1254] := 0.7489327;
   X[1255] := 0.841486;
   X[1256] := 0.944571;
   X[1257] := 1.047401;
   X[1258] := 1.1493956;
   X[1259] := 1.2461296;
   X[1260] := 1.3409435;
   X[1261] := 1.4471296;
   X[1262] := 1.5429435;
   X[1263] := 1.6451297;
   X[1264] := 1.7413158;
   X[1265] := 1.8395978;
   X[1266] := 1.9470446;
   X[1267] := 2.046316;
   X[1268] := 2.141688;
   X[1269] := 2.2395074;
   X[1270] := 2.3439596;
   X[1271] := 2.440784;
   X[1272] := 2.540598;
   X[1273] := 2.6418743;
   X[1274] := 2.7417786;
   X[1275] := 2.8391511;
   X[1276] := 2.9425128;
   X[1277] := 3.0404222;
   X[1278] := 3.1325235;
   X[1279] := 3.2412467;
   X[1280] := 3.3387947;
   X[1281] := 3.4342575;
   X[1282] := 3.5342574;
   X[1283] := 3.6396246;
   X[1284] := 3.7380767;
   X[1285] := 3.8398108;
   X[1286] := 3.9381723;
   X[1287] := 4.034534;
   X[1288] := 4.13063;
   X[1289] := 4.2379065;
   X[1290] := 4.332268;
   X[1291] := 4.4399066;
   X[1292] := 4.5368214;
   X[1293] := 4.628816;
   X[1294] := 4.735364;
   X[1295] := 4.836087;
   X[1296] := 4.928742;
   X[1297] := 5.0387416;
   X[1298] := 5.130109;
   X[1299] := 5.239098;
   X[1300] := 5.3370132;
   X[1301] := 5.43438;
   X[1302] := 5.5339227;
   X[1303] := 5.6311035;
   X[1304] := 5.731024;
   X[1305] := 5.8305664;
   X[1306] := 5.924747;
   X[1307] := 6.027933;
   X[1308] := 6.1294813;
   X[1309] := 6.2354865;
   X[1310] := 6.3234863;
   X[1311] := 6.43004;
   X[1312] := 6.530306;
   X[1313] := 6.6274014;
   X[1314] := 6.7249546;
   X[1315] := 6.8309493;
   X[1316] := 6.9234123;
   X[1317] := 7.0274973;
   X[1318] := 7.1264067;
   X[1319] := 7.2263165;
   X[1320] := 7.329322;
   X[1321] := 7.422141;
   X[1322] := 7.5283217;
   X[1323] := 7.6280613;
   X[1324] := 7.7241464;
   X[1325] := 7.820609;
   X[1326] := 7.923875;
   X[1327] := 8.022885;
   X[1328] := 8.123976;
   X[1329] := 8.231061;
   X[1330] := 8.323157;
   X[1331] := 8.426066;
   X[1332] := 8.522167;
   X[1333] := 8.62453;
   X[1334] := 8.719806;
   X[1335] := 8.822077;
   X[1336] := 8.918812;
   X[1337] := 9.018099;
   X[1338] := 9.116663;
   X[1339] := 9.21195;
   X[1340] := 9.308865;
   X[1341] := 9.403785;
   X[1342] := 9.504344;
   X[1343] := 9.603817;
   X[1344] := 9.694104;
   X[1345] := 9.796387;
   X[1346] := 9.90503;
   X[1347] := 9.994046;
   X[1348] := 10.088147;
   X[1349] := 10.185254;
   X[1350] := 10.283903;
   X[1351] := 10.380095;
   X[1352] := 10.480473;
   X[1353] := 10.572754;
   X[1354] := 10.679222;
   X[1355] := 10.772696;
   X[1356] := 10.870611;
   X[1357] := 10.970898;
   X[1358] := 11.067276;
   X[1359] := 11.16219;
   X[1360] := 11.261116;
   X[1361] := 11.365132;
   X[1362] := 11.458878;
   X[1363] := 11.550426;
   X[1364] := 11.658532;
   X[1365] := 11.751276;
   X[1366] := 11.844559;
   X[1367] := 11.944931;
   X[1368] := 12.048128;
   X[1369] := 12.144404;
   X[1370] := 12.240521;
   X[1371] := 12.341804;
   X[1372] := 12.436001;
   X[1373] := 12.537735;
   X[1374] := 12.632028;
   X[1375] := 12.722315;
   X[1376] := 12.822873;
   X[1377] := 12.918155;
   X[1378] := 13.020804;
   X[1379] := 13.11182;
   X[1380] := 13.215831;
   X[1381] := 13.312203;
   X[1382] := 13.411315;
   X[1383] := 13.506406;
   X[1384] := 13.602703;
   X[1385] := 13.704895;
   X[1386] := 13.813751;
   X[1387] := 13.936825;
   X[1388] := 14.052898;
   X[1389] := 14.177792;
   X[1390] := 14.293041;
   X[1391] := 14.399817;
   X[1392] := 14.500093;
   X[1393] := 14.601089;
   X[1394] := 14.699647;
   X[1395] := 14.798828;
   X[1396] := 14.900009;
   X[1397] := 14.99928;
   X[1398] := 15.095919;
   X[1399] := 15.194653;
   X[1400] := 15.2962055;
   X[1401] := 15.402014;
   X[1402] := 15.493297;
   X[1403] := 15.597206;
   X[1404] := 15.696291;
   X[1405] := 15.793211;
   X[1406] := 15.894573;
   X[1407] := 15.994216;
   X[1408] := 16.094482;
   X[1409] := 16.197584;
   X[1410] := 16.296854;
   X[1411] := 16.395493;
   X[1412] := 16.494854;
   X[1413] := 16.593866;
   X[1414] := 16.69186;
   X[1415] := 16.793776;
   X[1416] := 16.89269;
   X[1417] := 16.994047;
   X[1418] := 17.094774;
   X[1419] := 17.193243;
   X[1420] := 17.292328;
   X[1421] := 17.389967;
   X[1422] := 17.489605;
   X[1423] := 17.591696;
   X[1424] := 17.690153;
   X[1425] := 17.79379;
   X[1426] := 17.88644;
   X[1427] := 17.984615;
   X[1428] := 18.091429;
   X[1429] := 18.188078;
   X[1430] := 18.289797;
   X[1431] := 18.389711;
   X[1432] := 18.487074;
   X[1433] := 18.585089;
   X[1434] := 18.683716;
   X[1435] := 18.787716;
   X[1436] := 18.88736;
   X[1437] := 18.982813;
   X[1438] := 19.084908;
   X[1439] := 19.180637;
   X[1440] := 19.287733;
   X[1441] := 19.378914;
   X[1442] := 19.481653;
   X[1443] := 19.58519;
   X[1444] := 19.688015;
   X[1445] := 19.784105;
   X[1446] := 19.885105;
   X[1447] := 19.981941;
   X[1448] := 20.080477;
   X[1449] := 20.177025;
   X[1450] := 20.277748;
   X[1451] := 20.381495;
   X[1452] := 20.474669;
   X[1453] := 20.585121;
   X[1454] := 20.684946;
   X[1455] := 20.782211;
   X[1456] := 20.869228;
   X[1457] := 20.983856;
   X[1458] := 21.075409;
   X[1459] := 21.175041;
   X[1460] := 21.27759;
   X[1461] := 21.37559;
   X[1462] := 21.48168;
   X[1463] := 21.57587;
   X[1464] := 21.669786;
   X[1465] := 21.769611;
   X[1466] := 21.87778;
   X[1467] := 21.970972;
   X[1468] := 22.07425;
   X[1469] := 22.1737;
   X[1470] := 22.27034;
   X[1471] := 22.372978;
   X[1472] := 22.464525;
   X[1473] := 22.568436;
   X[1474] := 22.673801;
   X[1475] := 22.76935;
   X[1476] := 22.873451;
   X[1477] := 22.968447;
   X[1478] := 23.068174;
   X[1479] := 23.167181;
   X[1480] := 23.262638;
   X[1481] := 23.363457;
   X[1482] := 23.448547;
   X[1483] := 23.490519;
   X[1484] := 23.525759;
   X[1485] := 23.558645;
   X[1486] := 23.595072;
   X[1487] := 23.638952;
   X[1488] := 23.6792;
   X[1489] := 23.715626;
   X[1490] := 23.748682;
   X[1491] := 23.789104;
   X[1492] := 23.828627;
   X[1493] := 23.864237;
   X[1494] := 23.902477;
   X[1495] := 23.940363;
   X[1496] := 23.9459;
   X[1497] := 23.91903;
   X[1498] := 23.88006;
   X[1499] := 23.848814;
   X[1500] := 23.799929;
   X[1501] := 23.76615;
   X[1502] := 23.732264;
   X[1503] := 23.693836;
   X[1504] := 23.654856;
   X[1505] := 23.61289;
   X[1506] := 23.575373;
   X[1507] := 23.54095;
   X[1508] := 23.499975;
   X[1509] := 23.465818;
   X[1510] := 23.40177;
   X[1511] := 23.306679;
   X[1512] := 23.211945;
   X[1513] := 23.113216;
   X[1514] := 23.009312;
   X[1515] := 22.915482;
   X[1516] := 22.810843;
   X[1517] := 22.714844;
   X[1518] := 22.607939;
   X[1519] := 22.5082;
   X[1520] := 22.41111;
   X[1521] := 22.315023;
   X[1522] := 22.216562;
   X[1523] := 22.114561;
   X[1524] := 22.017641;
   X[1525] := 21.91356;
   X[1526] := 21.818556;
   X[1527] := 21.71846;
   X[1528] := 21.61546;
   X[1529] := 21.519827;
   X[1530] := 21.423178;
   X[1531] := 21.322727;
   X[1532] := 21.2219;
   X[1533] := 21.118635;
   X[1534] := 21.017353;
   X[1535] := 20.921162;
   X[1536] := 20.821173;
   X[1537] := 20.717806;
   X[1538] := 20.617353;
   X[1539] := 20.519167;
   X[1540] := 20.423529;
   X[1541] := 20.323885;
   X[1542] := 20.222248;
   X[1543] := 20.122982;
   X[1544] := 20.017609;
   X[1545] := 19.922152;
   X[1546] := 19.82279;
   X[1547] := 19.728874;
   X[1548] := 19.628683;
   X[1549] := 19.527231;
   X[1550] := 19.420507;
   X[1551] := 19.328598;
   X[1552] := 19.226055;
   X[1553] := 19.12614;
   X[1554] := 19.027859;
   X[1555] := 18.92413;
   X[1556] := 18.830034;
   X[1557] := 18.725492;
   X[1558] := 18.621853;
   X[1559] := 18.528305;
   X[1560] := 18.429848;
   X[1561] := 18.329391;
   X[1562] := 18.231758;
   X[1563] := 18.133385;
   X[1564] := 18.02812;
   X[1565] := 17.93539;
   X[1566] := 17.828562;
   X[1567] := 17.731556;
   X[1568] := 17.632019;
   X[1569] := 17.53247;
   X[1570] := 17.435652;
   X[1571] := 17.331741;
   X[1572] := 17.23164;
   X[1573] := 17.13119;
   X[1574] := 17.039188;
   X[1575] := 16.934822;
   X[1576] := 16.834013;
   X[1577] := 16.72946;
   X[1578] := 16.632635;
   X[1579] := 16.541449;
   X[1580] := 16.433624;
   X[1581] := 16.337263;
   X[1582] := 16.238619;
   X[1583] := 16.140078;
   X[1584] := 16.041264;
   X[1585] := 15.936167;
   X[1586] := 15.837439;
   X[1587] := 15.731354;
   X[1588] := 15.643433;
   X[1589] := 15.542253;
   X[1590] := 15.437524;
   X[1591] := 15.340157;
   X[1592] := 15.234438;
   X[1593] := 15.1426935;
   X[1594] := 15.038332;
   X[1595] := 14.945151;
   X[1596] := 14.839055;
   X[1597] := 14.736237;
   X[1598] := 14.64305;
   X[1599] := 14.54605;
   X[1600] := 14.445321;
   X[1601] := 14.343502;
   X[1602] := 14.241587;
   X[1603] := 14.14296;
   X[1604] := 14.043225;
   X[1605] := 13.940954;
   X[1606] := 13.848028;
   X[1607] := 13.748943;
   X[1608] := 13.649853;
   X[1609] := 13.5404005;
   X[1610] := 13.445395;
   X[1611] := 13.346565;
   X[1612] := 13.251119;
   X[1613] := 13.149114;
   X[1614] := 13.047938;
   X[1615] := 12.949023;
   X[1616] := 12.845475;
   X[1617] := 12.744108;
   X[1618] := 12.648922;
   X[1619] := 12.546831;
   X[1620] := 12.443922;
   X[1621] := 12.351374;
   X[1622] := 12.2532835;
   X[1623] := 12.144917;
   X[1624] := 12.04564;
   X[1625] := 11.948273;
   X[1626] := 11.850539;
   X[1627] := 11.755182;
   X[1628] := 11.652087;
   X[1629] := 11.552539;
   X[1630] := 11.4536295;
   X[1631] := 11.353901;
   X[1632] := 11.25381;
   X[1633] := 11.150906;
   X[1634] := 11.051443;
   X[1635] := 10.959076;
   X[1636] := 10.856342;
   X[1637] := 10.759076;
   X[1638] := 10.655523;
   X[1639] := 10.555251;
   X[1640] := 10.460879;
   X[1641] := 10.356331;
   X[1642] := 10.25497;
   X[1643] := 10.159789;
   X[1644] := 10.060602;
   X[1645] := 9.955512;
   X[1646] := 9.858231;
   X[1647] := 9.758411;
   X[1648] := 9.658512;
   X[1649] := 9.55823;
   X[1650] := 9.461773;
   X[1651] := 9.35714;
   X[1652] := 9.258135;
   X[1653] := 9.159677;
   X[1654] := 9.060767;
   X[1655] := 8.962858;
   X[1656] := 8.86222;
   X[1657] := 8.762124;
   X[1658] := 8.663587;
   X[1659] := 8.565485;
   X[1660] := 8.465938;
   X[1661] := 8.362666;
   X[1662] := 8.270204;
   X[1663] := 8.161209;
   X[1664] := 8.063927;
   X[1665] := 7.969384;
   X[1666] := 7.865379;
   X[1667] := 7.757927;
   X[1668] := 7.661746;
   X[1669] := 7.571554;
   X[1670] := 7.4681025;
   X[1671] := 7.373012;
   X[1672] := 7.262645;
   X[1673] := 7.166826;
   X[1674] := 7.067826;
   X[1675] := 6.965905;
   X[1676] := 6.872453;
   X[1677] := 6.765549;
   X[1678] := 6.6689053;
   X[1679] := 6.567815;
   X[1680] := 6.467815;
   X[1681] := 6.374448;
   X[1682] := 6.27481;
   X[1683] := 6.170256;
   X[1684] := 6.0742564;
   X[1685] := 5.970443;
   X[1686] := 5.867533;
   X[1687] := 5.775799;
   X[1688] := 5.669251;
   X[1689] := 5.576607;
   X[1690] := 5.4744263;
   X[1691] := 5.37507;
   X[1692] := 5.274251;
   X[1693] := 5.173602;
   X[1694] := 5.0736976;
   X[1695] := 4.973969;
   X[1696] := 4.87824;
   X[1697] := 4.7821445;
   X[1698] := 4.680597;
   X[1699] := 4.5706925;
   X[1700] := 4.4696817;
   X[1701] := 4.3800435;
   X[1702] := 4.268049;
   X[1703] := 4.172134;
   X[1704] := 4.080586;
   X[1705] := 3.9725008;
   X[1706] := 3.8796763;
   X[1707] := 3.7860382;
   X[1708] := 3.6812189;
   X[1709] := 3.5841231;
   X[1710] := 3.479304;
   X[1711] := 3.376038;
   X[1712] := 3.285123;
   X[1713] := 3.1766655;
   X[1714] := 3.0816603;
   X[1715] := 2.9889317;
   X[1716] := 2.8742027;
   X[1717] := 2.7805698;
   X[1718] := 2.6814742;
   X[1719] := 2.58474;
   X[1720] := 2.4808357;
   X[1721] := 2.3843784;
   X[1722] := 2.2894688;
   X[1723] := 2.1821017;
   X[1724] := 2.0858252;
   X[1725] := 1.9848198;
   X[1726] := 1.8824581;
   X[1727] := 1.7823783;
   X[1728] := 1.689091;
   X[1729] := 1.5809155;
   X[1730] := 1.4890857;
   X[1731] := 1.3824581;
   X[1732] := 1.2849952;
   X[1733] := 1.1856335;
   X[1734] := 1.0859048;
   X[1735] := 0.9898941;
   X[1736] := 0.8930803;
   X[1737] := 0.7830696;
   X[1738] := 0.6876282;
   X[1739] := 0.5891654;
   X[1740] := 0.48952705;
   X[1741] := 0.39324507;
   X[1742] := 0.29234084;
   X[1743] := 0.20517014;
   X[1744] := 0.11862703;
   X[1745] := 0.044536024;
   X[1747] := 0.059942853;
   X[1748] := 0.15758651;
   X[1749] := 0.25440568;
   X[1750] := 0.3589482;
   X[1751] := 0.46004933;
   X[1752] := 0.5611344;
   X[1753] := 0.6548631;
   X[1754] := 0.75676733;
   X[1755] := 0.86150146;
   X[1756] := 0.95358115;
   X[1757] := 1.0613099;
   X[1758] := 1.1569589;
   X[1759] := 1.2548631;
   X[1760] := 1.3582249;
   X[1761] := 1.4564961;
   X[1762] := 1.5571398;
   X[1763] := 1.6575068;
   X[1764] := 1.7561344;
   X[1765] := 1.8561398;
   X[1766] := 1.9555973;
   X[1767] := 2.055959;
   X[1768] := 2.15731;
   X[1769] := 2.2549536;
   X[1770] := 2.355693;
   X[1771] := 2.4565973;
   X[1772] := 2.5547833;
   X[1773] := 2.653778;
   X[1774] := 2.7529643;
   X[1775] := 2.8573205;
   X[1776] := 2.9499643;
   X[1777] := 3.0485973;
   X[1778] := 3.154326;
   X[1779] := 3.258145;
   X[1780] := 3.3519697;
   X[1781] := 3.4530602;
   X[1782] := 3.5616877;
   X[1783] := 3.6537888;
   X[1784] := 3.7530653;
   X[1785] := 3.8539696;
   X[1786] := 3.9496984;
   X[1787] := 4.048975;
   X[1788] := 4.15506;
   X[1789] := 4.2600656;
   X[1790] := 4.3559694;
   X[1791] := 4.450241;
   X[1792] := 4.553613;
   X[1793] := 4.6583314;
   X[1794] := 4.7553368;
   X[1795] := 4.8541613;
   X[1796] := 4.952624;
   X[1797] := 5.0506186;
   X[1798] := 5.1556134;
   X[1799] := 5.2568846;
   X[1800] := 5.3572516;
   X[1801] := 5.4571557;
   X[1802] := 5.5487146;
   X[1803] := 5.6542516;
   X[1804] := 5.7500815;
   X[1805] := 5.848257;
   X[1806] := 5.946342;
   X[1807] := 6.0442944;
   X[1808] := 6.131662;
   X[1809] := 6.2118382;
   X[1810] := 6.2960143;
   X[1811] := 6.375015;
   X[1812] := 6.475398;
   X[1813] := 6.5699406;
   X[1814] := 6.673946;
   X[1815] := 6.7746744;
   X[1816] := 6.876488;
   X[1817] := 6.9773183;
   X[1818] := 7.0665946;
   X[1819] := 7.1729617;
   X[1820] := 7.27168;
   X[1821] := 7.3722386;
   X[1822] := 7.4740577;
   X[1823] := 7.5736055;
   X[1824] := 7.6791425;
   X[1825] := 7.767797;
   X[1826] := 7.8653398;
   X[1827] := 7.969797;
   X[1828] := 8.065621;
   X[1829] := 8.167153;
   X[1830] := 8.269989;
   X[1831] := 8.361536;
   X[1832] := 8.461175;
   X[1833] := 8.568446;
   X[1834] := 8.663994;
   X[1835] := 8.763;
   X[1836] := 8.869728;
   X[1837] := 8.967185;
   X[1838] := 9.065;
   X[1839] := 9.166371;
   X[1840] := 9.254648;
   X[1841] := 9.360101;
   X[1842] := 9.46093;
   X[1843] := 9.563106;
   X[1844] := 9.661111;
   X[1845] := 9.7617445;
   X[1846] := 9.856659;
   X[1847] := 9.962297;
   X[1848] := 10.057298;
   X[1849] := 10.164111;
   X[1850] := 10.258941;
   X[1851] := 10.361484;
   X[1852] := 10.453223;
   X[1853] := 10.551409;
   X[1854] := 10.659042;
   X[1855] := 10.756239;
   X[1856] := 10.855047;
   X[1857] := 10.954414;
   X[1858] := 11.057234;
   X[1859] := 11.149872;
   X[1860] := 11.254872;
   X[1861] := 11.352612;
   X[1862] := 11.447612;
   X[1863] := 11.55634;
   X[1864] := 11.652515;
   X[1865] := 11.749978;
   X[1866] := 11.846899;
   X[1867] := 11.953888;
   X[1868] := 12.050718;
   X[1869] := 12.148436;
   X[1870] := 12.250532;
   X[1871] := 12.347176;
   X[1872] := 12.448813;
   X[1873] := 12.549452;
   X[1874] := 12.646452;
   X[1875] := 12.7430105;
   X[1876] := 12.8481865;
   X[1877] := 12.946457;
   X[1878] := 13.047372;
   X[1879] := 13.147378;
   X[1880] := 13.250473;
   X[1881] := 13.3443775;
   X[1882] := 13.441564;
   X[1883] := 13.545021;
   X[1884] := 13.642846;
   X[1885] := 13.746388;
   X[1886] := 13.845665;
   X[1887] := 13.943575;
   X[1888] := 14.038495;
   X[1889] := 14.137947;
   X[1890] := 14.241128;
   X[1891] := 14.341495;
   X[1892] := 14.437409;
   X[1893] := 14.545048;
   X[1894] := 14.636771;
   X[1895] := 14.736697;
   X[1896] := 14.835883;
   X[1897] := 14.933149;
   X[1898] := 15.03534;
   X[1899] := 15.131453;
   X[1900] := 15.23091;
   X[1901] := 15.330197;
   X[1902] := 15.4204;
   X[1903] := 15.52323;
   X[1904] := 15.6187935;
   X[1905] := 15.709166;
   X[1906] := 15.815352;
   X[1907] := 15.914922;
   X[1908] := 16.00639;
   X[1909] := 16.110039;
   X[1910] := 16.208954;
   X[1911] := 16.302608;
   X[1912] := 16.396261;
   X[1913] := 16.497183;
   X[1914] := 16.591007;
   X[1915] := 16.693203;
   X[1916] := 16.793215;
   X[1917] := 16.88896;
   X[1918] := 16.986065;
   X[1919] := 17.089806;
   X[1920] := 17.184998;
   X[1921] := 17.2752;
   X[1922] := 17.376476;
   X[1923] := 17.468401;
   X[1924] := 17.57196;
   X[1925] := 17.669874;
   X[1926] := 17.769077;
   X[1927] := 17.861189;
   X[1928] := 17.959019;
   X[1929] := 18.059114;
   X[1930] := 18.161945;
   X[1931] := 18.251875;
   X[1932] := 18.350977;
   X[1933] := 18.449902;
   X[1934] := 18.548456;
   X[1935] := 18.64293;
   X[1936] := 18.740578;
   X[1937] := 18.837872;
   X[1938] := 18.937328;
   X[1939] := 19.02971;
   X[1940] := 19.129723;
   X[1941] := 19.232094;
   X[1942] := 19.325014;
   X[1943] := 19.422764;
   X[1944] := 19.525595;
   X[1945] := 19.613792;
   X[1946] := 19.719078;
   X[1947] := 19.814;
   X[1948] := 19.919504;
   X[1949] := 20.04212;
   X[1950] := 20.15819;
   X[1951] := 20.281082;
   X[1952] := 20.401524;
   X[1953] := 20.511564;
   X[1954] := 20.60375;
   X[1955] := 20.707033;
   X[1956] := 20.808395;
   X[1957] := 20.91049;
   X[1958] := 21.010033;
   X[1959] := 21.10931;
   X[1960] := 21.2064;
   X[1961] := 21.304592;
   X[1962] := 21.406315;
   X[1963] := 21.508495;
   X[1964] := 21.6065;
   X[1965] := 21.704512;
   X[1966] := 21.798693;
   X[1967] := 21.906687;
   X[1968] := 21.997974;
   X[1969] := 22.100151;
   X[1970] := 22.204704;
   X[1971] := 22.302252;
   X[1972] := 22.39762;
   X[1973] := 22.504076;
   X[1974] := 22.600353;
   X[1975] := 22.696167;
   X[1976] := 22.79672;
   X[1977] := 22.903719;
   X[1978] := 22.993368;
   X[1979] := 23.094183;
   X[1980] := 23.198092;
   X[1981] := 23.299007;
   X[1982] := 23.396645;
   X[1983] := 23.495646;
   X[1984] := 23.593475;
   X[1985] := 23.692747;
   X[1986] := 23.791107;
   X[1987] := 23.893204;
   X[1988] := 23.99648;
   X[1989] := 24.092756;
   X[1990] := 24.191118;
   X[1991] := 24.289673;
   X[1992] := 24.395853;
   X[1993] := 24.491858;
   X[1994] := 24.584322;
   X[1995] := 24.686327;
   X[1996] := 24.790226;
   X[1997] := 24.88778;
   X[1998] := 24.98996;
   X[1999] := 25.084875;
   X[2000] := 25.183603;
   X[2001] := 25.28597;
   X[2002] := 25.391157;
   X[2003] := 25.48106;
   X[2004] := 25.583986;
   X[2005] := 25.681438;
   X[2006] := 25.78654;
   X[2007] := 25.882534;
   X[2008] := 25.976997;
   X[2009] := 26.084625;
   X[2010] := 26.178997;
   X[2011] := 26.279093;
   X[2012] := 26.380821;
   X[2013] := 26.480001;
   X[2014] := 26.584827;
   X[2015] := 26.674923;
   X[2016] := 26.775928;
   X[2017] := 26.882019;
   X[2018] := 26.97811;
   X[2019] := 27.076385;
   X[2020] := 27.172386;
   X[2021] := 27.27448;
   X[2022] := 27.374933;
   X[2023] := 27.473944;
   X[2024] := 27.57186;
   X[2025] := 27.674858;
   X[2026] := 27.774858;
   X[2027] := 27.871407;
   X[2028] := 27.970226;
   X[2029] := 28.07169;
   X[2030] := 28.170599;
   X[2031] := 28.272417;
   X[2032] := 28.366512;
   X[2033] := 28.4667;
   X[2034] := 28.564981;
   X[2035] := 28.665806;
   X[2036] := 28.770975;
   X[2037] := 28.865072;
   X[2038] := 28.963987;
   X[2039] := 29.059992;
   X[2040] := 29.169172;
   X[2041] := 29.265812;
   X[2042] := 29.362364;
   X[2043] := 29.462551;
   X[2044] := 29.55378;
   X[2045] := 29.593468;
   X[2046] := 29.635618;
   X[2047] := 29.666414;
   X[2048] := 29.698565;
   X[2049] := 29.740263;
   X[2050] := 29.778048;
   X[2051] := 29.8223;
   X[2052] := 29.86127;
   X[2053] := 29.90024;
   X[2054] := 29.936306;
   X[2055] := 29.971361;
   X[2056] := 29.971085;
   X[2057] := 29.944763;
   X[2058] := 29.909967;
   X[2059] := 29.872366;
   X[2060] := 29.835667;
   X[2061] := 29.80542;
   X[2062] := 29.759996;
   X[2063] := 29.717112;
   X[2064] := 29.685328;
   X[2065] := 29.645077;
   X[2066] := 29.608839;
   X[2067] := 29.573593;
   X[2068] := 29.501139;
   X[2069] := 29.405039;
   X[2070] := 29.305681;
   X[2071] := 29.206215;
   X[2072] := 29.103575;
   X[2073] := 29.009033;
   X[2074] := 28.904667;
   X[2075] := 28.804937;
   X[2076] := 28.710293;
   X[2077] := 28.605474;
   X[2078] := 28.508661;
   X[2079] := 28.417282;
   X[2080] := 28.311565;
   X[2081] := 28.214464;
   X[2082] := 28.114277;
   X[2083] := 28.012548;
   X[2084] := 27.913092;
   X[2085] := 27.820448;
   X[2086] := 27.71899;
   X[2087] := 27.618353;
   X[2088] := 27.514618;
   X[2089] := 27.415438;
   X[2090] := 27.320534;
   X[2091] := 27.218431;
   X[2092] := 27.11598;
   X[2093] := 27.018234;
   X[2094] := 26.922245;
   X[2095] := 26.822065;
   X[2096] := 26.722776;
   X[2097] := 26.62123;
   X[2098] := 26.523596;
   X[2099] := 26.426495;
   X[2100] := 26.323044;
   X[2101] := 26.222862;
   X[2102] := 26.12549;
   X[2103] := 26.024942;
   X[2104] := 25.92758;
   X[2105] := 25.820772;
   X[2106] := 25.725574;
   X[2107] := 25.629202;
   X[2108] := 25.528017;
   X[2109] := 25.425926;
   X[2110] := 25.324293;
   X[2111] := 25.22792;
   X[2112] := 25.126825;
   X[2113] := 25.029005;
   X[2114] := 24.933367;
   X[2115] := 24.829548;
   X[2116] := 24.730543;
   X[2117] := 24.63091;
   X[2118] := 24.531271;
   X[2119] := 24.427984;
   X[2120] := 24.337261;
   X[2121] := 24.231985;
   X[2122] := 24.136707;
   X[2123] := 24.031889;
   X[2124] := 23.931883;
   X[2125] := 23.831882;
   X[2126] := 23.73997;
   X[2127] := 23.641516;
   X[2128] := 23.532425;
   X[2129] := 23.435963;
   X[2130] := 23.343596;
   X[2131] := 23.237778;
   X[2132] := 23.142862;
   X[2133] := 23.039133;
   X[2134] := 22.941957;
   X[2135] := 22.839037;
   X[2136] := 22.74458;
   X[2137] := 22.63958;
   X[2138] := 22.542213;
   X[2139] := 22.444937;
   X[2140] := 22.347937;
   X[2141] := 22.243298;
   X[2142] := 22.14175;
   X[2143] := 22.049746;
   X[2144] := 21.94365;
   X[2145] := 21.849377;
   X[2146] := 21.7401;
   X[2147] := 21.650915;
   X[2148] := 21.54883;
   X[2149] := 21.443733;
   X[2150] := 21.34736;
   X[2151] := 21.248903;
   X[2152] := 21.14999;
   X[2153] := 21.053713;
   X[2154] := 20.948261;
   X[2155] := 20.850527;
   X[2156] := 20.752527;
   X[2157] := 20.654068;
   X[2158] := 20.551973;
   X[2159] := 20.450611;
   X[2160] := 20.353426;
   X[2161] := 20.247616;
   X[2162] := 20.158962;
   X[2163] := 20.056686;
   X[2164] := 19.95451;
   X[2165] := 19.848787;
   X[2166] := 19.76441;
   X[2167] := 19.6565;
   X[2168] := 19.555319;
   X[2169] := 19.45823;
   X[2170] := 19.358404;
   X[2171] := 19.264393;
   X[2172] := 19.158207;
   X[2173] := 19.05784;
   X[2174] := 18.959488;
   X[2175] := 18.859291;
   X[2176] := 18.76084;
   X[2177] := 18.65584;
   X[2178] := 18.561293;
   X[2179] := 18.458387;
   X[2180] := 18.365738;
   X[2181] := 18.261276;
   X[2182] := 18.16474;
   X[2183] := 18.065456;
   X[2184] := 17.959185;
   X[2185] := 17.868;
   X[2186] := 17.770355;
   X[2187] := 17.661999;
   X[2188] := 17.565441;
   X[2189] := 17.466255;
   X[2190] := 17.363897;
   X[2191] := 17.270435;
   X[2192] := 17.170887;
   X[2193] := 17.071249;
   X[2194] := 16.968435;
   X[2195] := 16.872057;
   X[2196] := 16.771149;
   X[2197] := 16.675966;
   X[2198] := 16.571058;
   X[2199] := 16.47269;
   X[2200] := 16.371775;
   X[2201] := 16.271776;
   X[2202] := 16.172047;
   X[2203] := 16.071234;
   X[2204] := 15.967866;
   X[2205] := 15.878132;
   X[2206] := 15.776042;
   X[2207] := 15.676312;
   X[2208] := 15.57985;
   X[2209] := 15.473297;
   X[2210] := 15.378382;
   X[2211] := 15.279025;
   X[2212] := 15.177201;
   X[2213] := 15.079201;
   X[2214] := 14.981653;
   X[2215] := 14.875744;
   X[2216] := 14.789733;
   X[2217] := 14.678914;
   X[2218] := 14.583095;
   X[2219] := 14.475462;
   X[2220] := 14.384275;
   X[2221] := 14.279727;
   X[2222] := 14.186456;
   X[2223] := 14.079722;
   X[2224] := 13.987535;
   X[2225] := 13.88844;
   X[2226] := 13.783078;
   X[2227] := 13.69144;
   X[2228] := 13.58844;
   X[2229] := 13.489435;
   X[2230] := 13.387791;
   X[2231] := 13.282164;
   X[2232] := 13.192785;
   X[2233] := 13.088605;
   X[2234] := 12.986334;
   X[2235] := 12.884238;
   X[2236] := 12.789509;
   X[2237] := 12.687323;
   X[2238] := 12.587961;
   X[2239] := 12.48569;
   X[2240] := 12.391137;
   X[2241] := 12.28995;
   X[2242] := 12.1933975;
   X[2243] := 12.090126;
   X[2244] := 11.99194;
   X[2245] := 11.893216;
   X[2246] := 11.788483;
   X[2247] := 11.695754;
   X[2248] := 11.591849;
   X[2249] := 11.499387;
   X[2250] := 11.3926525;
   X[2251] := 11.294375;
   X[2252] := 11.194839;
   X[2253] := 11.092557;
   X[2254] := 10.997738;
   X[2255] := 10.890556;
   X[2256] := 10.798822;
   X[2257] := 10.69428;
   X[2258] := 10.595455;
   X[2259] := 10.501907;
   X[2260] := 10.401269;
   X[2261] := 10.301546;
   X[2262] := 10.204168;
   X[2263] := 10.10453;
   X[2264] := 9.9986315;
   X[2265] := 9.900072;
   X[2266] := 9.803525;
   X[2267] := 9.699344;
   X[2268] := 9.605338;
   X[2269] := 9.499519;
   X[2270] := 9.406876;
   X[2271] := 9.300428;
   X[2272] := 9.201333;
   X[2273] := 9.105418;
   X[2274] := 9.001323;
   X[2275] := 8.907136;
   X[2276] := 8.802052;
   X[2277] := 8.707588;
   X[2278] := 8.607865;
   X[2279] := 8.513311;
   X[2280] := 8.412035;
   X[2281] := 8.308216;
   X[2282] := 8.204583;
   X[2283] := 8.110939;
   X[2284] := 8.007684;
   X[2285] := 7.9073915;
   X[2286] := 7.813301;
   X[2287] := 7.709386;
   X[2288] := 7.6157475;
   X[2289] := 7.509753;
   X[2290] := 7.409833;
   X[2291] := 7.307189;
   X[2292] := 7.2156467;
   X[2293] := 7.115641;
   X[2294] := 7.0119123;
   X[2295] := 6.9109178;
   X[2296] := 6.8138165;
   X[2297] := 6.7170825;
   X[2298] := 6.618269;
   X[2299] := 6.5197263;
   X[2300] := 6.416269;
   X[2301] := 6.3316565;
   X[2302] := 6.241204;
   X[2303] := 6.1591926;
   X[2304] := 6.0856547;
   X[2305] := 5.9944844;
   X[2306] := 5.894399;
   X[2307] := 5.7966704;
   X[2308] := 5.6911173;
   X[2309] := 5.593761;
   X[2310] := 5.493942;
   X[2311] := 5.3995748;
   X[2312] := 5.2914844;
   X[2313] := 5.1911173;
   X[2314] := 5.095665;
   X[2315] := 4.987128;
   X[2316] := 4.8909416;
   X[2317] := 4.793027;
   X[2318] := 4.6963882;
   X[2319] := 4.5995693;
   X[2320] := 4.4999366;
   X[2321] := 4.4001174;
   X[2322] := 4.2952023;
   X[2323] := 4.1964736;
   X[2324] := 4.096298;
   X[2325] := 4.002112;
   X[2326] := 3.892383;
   X[2327] := 3.7965639;
   X[2328] := 3.6973832;
   X[2329] := 3.596197;
   X[2330] := 3.495383;
   X[2331] := 3.3942926;
   X[2332] := 3.2942874;
   X[2333] := 3.1958299;
   X[2334] := 3.094931;
   X[2335] := 2.997197;
   X[2336] := 2.8948298;
   X[2337] := 2.7965586;
   X[2338] := 2.6989202;
   X[2339] := 2.597463;
   X[2340] := 2.494101;
   X[2341] := 2.3953724;
   X[2342] := 2.299649;
   X[2343] := 2.196016;
   X[2344] := 2.1035533;
   X[2345] := 2.0005586;
   X[2346] := 1.9009149;
   X[2347] := 1.7969257;
   X[2348] := 1.702282;
   X[2349] := 1.5964628;
   X[2350] := 1.5001011;
   X[2351] := 1.3938245;
   X[2352] := 1.3030107;
   X[2353] := 1.1989149;
   X[2354] := 1.0978192;
   X[2355] := 0.99527663;
   X[2356] := 0.89845747;
   X[2357] := 0.8009096;
   X[2358] := 0.6996383;
   X[2359] := 0.60026056;
   X[2360] := 0.50273407;
   X[2361] := 0.39791492;
   X[2362] := 0.29663295;
   X[2363] := 0.20254253;
   X[2364] := 0.10845211;
   X[2365] := -0.0033723959;
   X[2367] := 0.025911892;
   X[2368] := 0.12764062;
   X[2369] := 0.2301778;
   X[2370] := 0.32582146;
   X[2371] := 0.42782146;
   X[2372] := 0.5292682;
   X[2373] := 0.6247364;
   X[2374] := 0.7245502;
   X[2375] := 0.82582146;
   X[2376] := 0.9259119;
   X[2377] := 1.0321778;
   X[2378] := 1.1327311;
   X[2379] := 1.2300928;
   X[2380] := 1.3288268;
   X[2381] := 1.4261938;
   X[2382] := 1.524731;
   X[2383] := 1.6241832;
   X[2384] := 1.7260131;
   X[2385] := 1.8231034;
   X[2386] := 1.9323747;
   X[2387] := 2.026098;
   X[2388] := 2.1261885;
   X[2389] := 2.2300076;
   X[2390] := 2.326013;
   X[2391] := 2.429545;
   X[2392] := 2.5251832;
   X[2393] := 2.626465;
   X[2394] := 2.7291992;
   X[2395] := 2.82646;
   X[2396] := 2.9284651;
   X[2397] := 3.0237417;
   X[2398] := 3.1271088;
   X[2399] := 3.2188323;
   X[2400] := 3.3277419;
   X[2401] := 3.4281034;
   X[2402] := 3.5262842;
   X[2403] := 3.6254652;
   X[2404] := 3.7312844;
   X[2405] := 3.8243802;
   X[2406] := 3.9309225;
   X[2407] := 4.0269175;
   X[2408] := 4.123109;
   X[2409] := 4.223928;
   X[2410] := 4.3228374;
   X[2411] := 4.425109;
   X[2412] := 4.525572;
   X[2413] := 4.6247525;
   X[2414] := 4.7195716;
   X[2415] := 4.822114;
   X[2416] := 4.9290237;
   X[2417] := 5.0293;
   X[2418] := 5.1238375;
   X[2419] := 5.2208376;
   X[2420] := 5.3288484;
   X[2421] := 5.4212046;
   X[2422] := 5.5208535;
   X[2423] := 5.6197524;
   X[2424] := 5.7191143;
   X[2425] := 5.8213906;
   X[2426] := 5.91721;
   X[2427] := 6.024593;
   X[2428] := 6.099498;
   X[2429] := 6.184956;
   X[2430] := 6.2723126;
   X[2431] := 6.350122;
   X[2432] := 6.4428988;
   X[2433] := 6.5479894;
   X[2434] := 6.6529894;
   X[2435] := 6.745814;
   X[2436] := 6.8487177;
   X[2437] := 6.9472713;
   X[2438] := 7.035271;
   X[2439] := 7.144271;
   X[2440] := 7.238819;
   X[2441] := 7.341181;
   X[2442] := 7.4426327;
   X[2443] := 7.544372;
   X[2444] := 7.642824;
   X[2445] := 7.739106;
   X[2446] := 7.842649;
   X[2447] := 7.943654;
   X[2448] := 8.03675;
   X[2449] := 8.132574;
   X[2450] := 8.232659;
   X[2451] := 8.330755;
   X[2452] := 8.439484;
   X[2453] := 8.538937;
   X[2454] := 8.632404;
   X[2455] := 8.740123;
   X[2456] := 8.838304;
   X[2457] := 8.93659;
   X[2458] := 9.036857;
   X[2459] := 9.1335;
   X[2460] := 9.236138;
   X[2461] := 9.329867;
   X[2462] := 9.441229;
   X[2463] := 9.532867;
   X[2464] := 9.63041;
   X[2465] := 9.731968;
   X[2466] := 9.836782;
   X[2467] := 9.934687;
   X[2468] := 10.030703;
   X[2469] := 10.1319685;
   X[2470] := 10.225612;
   X[2471] := 10.330792;
   X[2472] := 10.433166;
   X[2473] := 10.529888;
   X[2474] := 10.630798;
   X[2475] := 10.730081;
   X[2476] := 10.825798;
   X[2477] := 10.926899;
   X[2478] := 11.02517;
   X[2479] := 11.123815;
   X[2480] := 11.225634;
   X[2481] := 11.326186;
   X[2482] := 11.426543;
   X[2483] := 11.529186;
   X[2484] := 11.621825;
   X[2485] := 11.720729;
   X[2486] := 11.820463;
   X[2487] := 11.919373;
   X[2488] := 12.023655;
   X[2489] := 12.127926;
   X[2490] := 12.2206545;
   X[2491] := 12.318564;
   X[2492] := 12.427474;
   X[2493] := 12.514117;
   X[2494] := 12.62366;
   X[2495] := 12.719671;
   X[2496] := 12.820032;
   X[2497] := 12.917038;
   X[2498] := 13.015592;
   X[2499] := 13.123953;
   X[2500] := 13.222676;
   X[2501] := 13.317947;
   X[2502] := 13.420511;
   X[2503] := 13.5199585;
   X[2504] := 13.618325;
   X[2505] := 13.716778;
   X[2506] := 13.815873;
   X[2507] := 13.913511;
   X[2508] := 14.017325;
   X[2509] := 14.120155;
   X[2510] := 14.219336;
   X[2511] := 14.318698;
   X[2512] := 14.4135275;
   X[2513] := 14.515794;
   X[2514] := 14.611895;
   X[2515] := 14.711171;
   X[2516] := 14.814623;
   X[2517] := 14.910176;
   X[2518] := 15.008724;
   X[2519] := 15.108283;
   X[2520] := 15.208299;
   X[2521] := 15.299219;
   X[2522] := 15.397868;
   X[2523] := 15.499246;
   X[2524] := 15.597528;
   X[2525] := 15.69463;
   X[2526] := 15.784826;
   X[2527] := 15.888932;
   X[2528] := 15.987401;
   X[2529] := 16.084778;
   X[2530] := 16.17688;
   X[2531] := 16.277077;
   X[2532] := 16.375822;
   X[2533] := 16.474646;
   X[2534] := 16.573385;
   X[2535] := 16.667673;
   X[2536] := 16.769327;
   X[2537] := 16.866146;
   X[2538] := 16.960077;
   X[2539] := 17.057093;
   X[2540] := 17.158833;
   X[2541] := 17.259024;
   X[2542] := 17.352764;
   X[2543] := 17.458775;
   X[2544] := 17.544249;
   X[2545] := 17.644077;
   X[2546] := 17.743546;
   X[2547] := 17.84147;
   X[2548] := 17.936115;
   X[2549] := 18.032679;
   X[2550] := 18.130865;
   X[2551] := 18.22634;
   X[2552] := 18.327354;
   X[2553] := 18.425455;
   X[2554] := 18.527014;
   X[2555] := 18.623207;
   X[2556] := 18.719685;
   X[2557] := 18.813051;
   X[2558] := 18.916706;
   X[2559] := 19.010988;
   X[2560] := 19.104372;
   X[2561] := 19.19511;
   X[2562] := 19.297031;
   X[2563] := 19.396318;
   X[2564] := 19.499786;
   X[2565] := 19.601984;
   X[2566] := 19.691265;
   X[2567] := 19.786457;
   X[2568] := 19.895712;
   X[2569] := 20.013876;
   X[2570] := 20.135775;
   X[2571] := 20.25421;
   X[2572] := 20.382725;
   X[2573] := 20.4863;
   X[2574] := 20.591118;
   X[2575] := 20.683401;
   X[2576] := 20.788671;
   X[2577] := 20.885853;
   X[2578] := 20.984491;
   X[2579] := 21.08622;
   X[2580] := 21.181225;
   X[2581] := 21.282236;
   X[2582] := 21.384502;
   X[2583] := 21.48114;
   X[2584] := 21.588694;
   X[2585] := 21.678518;
   X[2586] := 21.781065;
   X[2587] := 21.880337;
   X[2588] := 21.975891;
   X[2589] := 22.07916;
   X[2590] := 22.182253;
   X[2591] := 22.2738;
   X[2592] := 22.384077;
   X[2593] := 22.48172;
   X[2594] := 22.582172;
   X[2595] := 22.679268;
   X[2596] := 22.774448;
   X[2597] := 22.880901;
   X[2598] := 22.972816;
   X[2599] := 23.07282;
   X[2600] := 23.175104;
   X[2601] := 23.271093;
   X[2602] := 23.370188;
   X[2603] := 23.478651;
   X[2604] := 23.57511;
   X[2605] := 23.670933;
   X[2606] := 23.773375;
   X[2607] := 23.874746;
   X[2608] := 23.974922;
   X[2609] := 24.07039;
   X[2610] := 24.167843;
   X[2611] := 24.270939;
   X[2612] := 24.375843;
   X[2613] := 24.473125;
   X[2614] := 24.571033;
   X[2615] := 24.666588;
   X[2616] := 24.763412;
   X[2617] := 24.86614;
   X[2618] := 24.969322;
   X[2619] := 25.059864;
   X[2620] := 25.162874;
   X[2621] := 25.268332;
   X[2622] := 25.369146;
   X[2623] := 25.4637;
   X[2624] := 25.556253;
   X[2625] := 25.663433;
   X[2626] := 25.759253;
   X[2627] := 25.857885;
   X[2628] := 25.96253;
   X[2629] := 26.060162;
   X[2630] := 26.153727;
   X[2631] := 26.260992;
   X[2632] := 26.36054;
   X[2633] := 26.461449;
   X[2634] := 26.56745;
   X[2635] := 26.662998;
   X[2636] := 26.755919;
   X[2637] := 26.854195;
   X[2638] := 26.961098;
   X[2639] := 27.058743;
   X[2640] := 27.158104;
   X[2641] := 27.25302;
   X[2642] := 27.356295;
   X[2643] := 27.460752;
   X[2644] := 27.554663;
   X[2645] := 27.651747;
   X[2646] := 27.752583;
   X[2647] := 27.850763;
   X[2648] := 27.956583;
   X[2649] := 28.05231;
   X[2650] := 28.153673;
   X[2651] := 28.251131;
   X[2652] := 28.347227;
   X[2653] := 28.45305;
   X[2654] := 28.550322;
   X[2655] := 28.644514;
   X[2656] := 28.746424;
   X[2657] := 28.850885;
   X[2658] := 28.945429;
   X[2659] := 29.045786;
   X[2660] := 29.144157;
   X[2661] := 29.248976;
   X[2662] := 29.344795;
   X[2663] := 29.447987;
   X[2664] := 29.54119;
   X[2665] := 29.580042;
   X[2666] := 29.62329;
   X[2667] := 29.656717;
   X[2668] := 29.69505;
   X[2669] := 29.733934;
   X[2670] := 29.772356;
   X[2671] := 29.803427;
   X[2672] := 29.852116;
   X[2673] := 29.881182;
   X[2674] := 29.923882;
   X[2675] := 29.96567;
   X[2676] := 29.996645;
   X[2677] := 29.996737;
   X[2678] := 29.976862;
   X[2679] := 29.937529;
   X[2680] := 29.899372;
   X[2681] := 29.862036;
   X[2682] := 29.82715;
   X[2683] := 29.790722;
   X[2684] := 29.751476;
   X[2685] := 29.716873;
   X[2686] := 29.671541;
   X[2687] := 29.637661;
   X[2688] := 29.600325;
   X[2689] := 29.562891;
   X[2690] := 29.493938;
   X[2691] := 29.387024;
   X[2692] := 29.2883;
   X[2693] := 29.18838;
   X[2694] := 29.090826;
   X[2695] := 28.990469;
   X[2696] := 28.890465;
   X[2697] := 28.78956;
   X[2698] := 28.687284;
   X[2699] := 28.590454;
   X[2700] := 28.49291;
   X[2701] := 28.390278;
   X[2702] := 28.291086;
   X[2703] := 28.196081;
   X[2704] := 28.096172;
   X[2705] := 27.991726;
   X[2706] := 27.88872;
   X[2707] := 27.7918;
   X[2708] := 27.692528;
   X[2709] := 27.598162;
   X[2710] := 27.50016;
   X[2711] := 27.389433;
   X[2712] := 27.29598;
   X[2713] := 27.19614;
   X[2714] := 27.10115;
   X[2715] := 26.999146;
   X[2716] := 26.898874;
   X[2717] := 26.802326;
   X[2718] := 26.699778;
   X[2719] := 26.604502;
   X[2720] := 26.505587;
   X[2721] := 26.398949;
   X[2722] := 26.30531;
   X[2723] := 26.21257;
   X[2724] := 26.1043;
   X[2725] := 26.00357;
   X[2726] := 25.900293;
   X[2727] := 25.804028;
   X[2728] := 25.70066;
   X[2729] := 25.603289;
   X[2730] := 25.501745;
   X[2731] := 25.402836;
   X[2732] := 25.309374;
   X[2733] := 25.207277;
   X[2734] := 25.106554;
   X[2735] := 25.017906;
   X[2736] := 24.908;
   X[2737] := 24.813635;
   X[2738] := 24.711176;
   X[2739] := 24.607452;
   X[2740] := 24.511442;
   X[2741] := 24.411905;
   X[2742] := 24.309532;
   X[2743] := 24.210623;
   X[2744] := 24.106895;
   X[2745] := 24.011885;
   X[2746] := 23.915064;
   X[2747] := 23.817879;
   X[2748] := 23.718336;
   X[2749] := 23.612879;
   X[2750] := 23.512873;
   X[2751] := 23.41915;
   X[2752] := 23.316235;
   X[2753] := 23.218868;
   X[2754] := 23.11732;
   X[2755] := 23.018139;
   X[2756] := 22.920315;
   X[2757] := 22.81941;
   X[2758] := 22.722948;
   X[2759] := 22.620123;
   X[2760] := 22.517574;
   X[2761] := 22.420574;
   X[2762] := 22.315123;
   X[2763] := 22.222755;
   X[2764] := 22.12566;
   X[2765] := 22.023117;
   X[2766] := 21.925192;
   X[2767] := 21.825563;
   X[2768] := 21.73065;
   X[2769] := 21.628372;
   X[2770] := 21.526367;
   X[2771] := 21.430271;
   X[2772] := 21.318914;
   X[2773] := 21.221;
   X[2774] := 21.128363;
   X[2775] := 21.02709;
   X[2776] := 20.929272;
   X[2777] := 20.824905;
   X[2778] := 20.726627;
   X[2779] := 20.62608;
   X[2780] := 20.528803;
   X[2781] := 20.428804;
   X[2782] := 20.329521;
   X[2783] := 20.232985;
   X[2784] := 20.126698;
   X[2785] := 20.030516;
   X[2786] := 19.936245;
   X[2787] := 19.833143;
   X[2788] := 19.73016;
   X[2789] := 19.634686;
   X[2790] := 19.531963;
   X[2791] := 19.437681;
   X[2792] := 19.332415;
   X[2793] := 19.23041;
   X[2794] := 19.130772;
   X[2795] := 19.034128;
   X[2796] := 18.935862;
   X[2797] := 18.835857;
   X[2798] := 18.7344;
   X[2799] := 18.637123;
   X[2800] := 18.539303;
   X[2801] := 18.435846;
   X[2802] := 18.342299;
   X[2803] := 18.23548;
   X[2804] := 18.132648;
   X[2805] := 18.038568;
   X[2806] := 17.937197;
   X[2807] := 17.84265;
   X[2808] := 17.740011;
   X[2809] := 17.6401;
   X[2810] := 17.539553;
   X[2811] := 17.443005;
   X[2812] := 17.345728;
   X[2813] := 17.248362;
   X[2814] := 17.139723;
   X[2815] := 17.042265;
   X[2816] := 16.949175;
   X[2817] := 16.84508;
   X[2818] := 16.7459;
   X[2819] := 16.651165;
   X[2820] := 16.548887;
   X[2821] := 16.443527;
   X[2822] := 16.346441;
   X[2823] := 16.250431;
   X[2824] := 16.14734;
   X[2825] := 16.052414;
   X[2826] := 15.950516;
   X[2827] := 15.8478775;
   X[2828] := 15.748414;
   X[2829] := 15.6508665;
   X[2830] := 15.549968;
   X[2831] := 15.453686;
   X[2832] := 15.353233;
   X[2833] := 15.2566805;
   X[2834] := 15.15468;
   X[2835] := 15.050313;
   X[2836] := 14.949765;
   X[2837] := 14.850856;
   X[2838] := 14.756941;
   X[2839] := 14.651936;
   X[2840] := 14.55458;
   X[2841] := 14.456659;
   X[2842] := 14.354032;
   X[2843] := 14.254026;
   X[2844] := 14.164557;
   X[2845] := 14.057015;
   X[2846] := 13.9621;
   X[2847] := 13.859839;
   X[2848] := 13.757015;
   X[2849] := 13.659914;
   X[2850] := 13.562005;
   X[2851] := 13.460457;
   X[2852] := 13.358547;
   X[2853] := 13.261728;
   X[2854] := 13.160632;
   X[2855] := 13.05718;
   X[2856] := 12.960356;
   X[2857] := 12.859446;
   X[2858] := 12.753175;
   X[2859] := 12.659808;
   X[2860] := 12.562978;
   X[2861] := 12.462707;
   X[2862] := 12.362706;
   X[2863] := 12.260882;
   X[2864] := 12.162425;
   X[2865] := 12.066069;
   X[2866] := 11.965696;
   X[2867] := 11.861158;
   X[2868] := 11.766967;
   X[2869] := 11.663696;
   X[2870] := 11.5686;
   X[2871] := 11.47168;
   X[2872] := 11.362696;
   X[2873] := 11.268866;
   X[2874] := 11.17177;
   X[2875] := 11.066137;
   X[2876] := 10.965228;
   X[2877] := 10.866946;
   X[2878] := 10.769228;
   X[2879] := 10.670036;
   X[2880] := 10.572036;
   X[2881] := 10.473488;
   X[2882] := 10.372393;
   X[2883] := 10.273207;
   X[2884] := 10.173297;
   X[2885] := 10.077653;
   X[2886] := 9.974563;
   X[2887] := 9.869749;
   X[2888] := 9.773738;
   X[2889] := 9.665658;
   X[2890] := 9.570834;
   X[2891] := 9.477557;
   X[2892] := 9.377461;
   X[2893] := 9.272547;
   X[2894] := 9.181094;
   X[2895] := 9.080542;
   X[2896] := 8.974089;
   X[2897] := 8.876733;
   X[2898] := 8.78218;
   X[2899] := 8.680536;
   X[2900] := 8.580536;
   X[2901] := 8.477078;
   X[2902] := 8.378435;
   X[2903] := 8.278711;
   X[2904] := 8.181706;
   X[2905] := 8.077887;
   X[2906] := 7.98052;
   X[2907] := 7.883791;
   X[2908] := 7.7804294;
   X[2909] := 7.676073;
   X[2910] := 7.583424;
   X[2911] := 7.4855146;
   X[2912] := 7.3815036;
   X[2913] := 7.286509;
   X[2914] := 7.1853228;
   X[2915] := 7.087509;
   X[2916] := 6.980594;
   X[2917] := 6.885408;
   X[2918] := 6.786227;
   X[2919] := 6.686775;
   X[2920] := 6.5914025;
   X[2921] := 6.4840407;
   X[2922] := 6.388397;
   X[2923] := 6.300397;
   X[2924] := 6.2213163;
   X[2925] := 6.139406;
   X[2926] := 6.047693;
   X[2927] := 5.965804;
   X[2928] := 5.8651657;
   X[2929] := 5.7661657;
   X[2930] := 5.66598;
   X[2931] := 5.567799;
   X[2932] := 5.463437;
   X[2933] := 5.359437;
   X[2934] := 5.2632565;
   X[2935] := 5.167432;
   X[2936] := 5.0657086;
   X[2937] := 4.9659796;
   X[2938] := 4.869437;
   X[2939] := 4.767799;
   X[2940] := 4.6630754;
   X[2941] := 4.566336;
   X[2942] := 4.463347;
   X[2943] := 4.3684425;
   X[2944] := 4.268799;
   X[2945] := 4.167703;
   X[2946] := 4.0643415;
   X[2947] := 3.9627085;
   X[2948] := 3.866432;
   X[2949] := 3.765517;
   X[2950] := 3.666788;
   X[2951] := 3.5658894;
   X[2952] := 3.468703;
   X[2953] := 3.3619797;
   X[2954] := 3.2612457;
   X[2955] := 3.1599743;
   X[2956] := 3.0651553;
   X[2957] := 2.9675224;
   X[2958] := 2.867517;
   X[2959] := 2.7654264;
   X[2960] := 2.6686072;
   X[2961] := 2.567969;
   X[2962] := 2.4646127;
   X[2963] := 2.3662403;
   X[2964] := 2.2672458;
   X[2965] := 2.1639743;
   X[2966] := 2.0745115;
   X[2967] := 1.9656924;
   X[2968] := 1.8648787;
   X[2969] := 1.7657936;
   X[2970] := 1.6727935;
   X[2971] := 1.5732456;
   X[2972] := 1.4724212;
   X[2973] := 1.3685116;
   X[2974] := 1.2602403;
   X[2975] := 1.1676978;
   X[2976] := 1.0685116;
   X[2977] := 0.97042114;
   X[2978] := 0.8631499;
   X[2979] := 0.77142113;
   X[2980] := 0.6708733;
   X[2981] := 0.5715966;
   X[2982] := 0.4670541;
   X[2983] := 0.36605412;
   X[2984] := 0.26659665;
   X[2985] := 0.16896369;
   X[2986] := 0.065697774;
   X[2987] := 0.04820052;
   X[2989] := -0.0073742764;
   X[2990] := 0.030601272;
   X[2991] := 0.12714916;
   X[2992] := 0.23242578;
   X[2993] := 0.33032465;
   X[2994] := 0.42942578;
   X[2995] := 0.532697;
   X[2996] := 0.63269705;
   X[2997] := 0.7281492;
   X[2998] := 0.8335109;
   X[2999] := 0.93724495;
   X[3000] := 1.0296971;
   X[3001] := 1.1316066;
   X[3002] := 1.2371545;
   X[3003] := 1.3257928;
   X[3004] := 1.4277024;
   X[3005] := 1.5306174;
   X[3006] := 1.6274258;
   X[3007] := 1.7276067;
   X[3008] := 1.8318886;
   X[3009] := 1.9328833;
   X[3010] := 2.0303407;
   X[3011] := 2.1277025;
   X[3012] := 2.2318885;
   X[3013] := 2.3308885;
   X[3014] := 2.4322503;
   X[3015] := 2.535878;
   X[3016] := 2.6287982;
   X[3017] := 2.726346;
   X[3018] := 2.8281653;
   X[3019] := 2.9279845;
   X[3020] := 3.0230694;
   X[3021] := 3.1296172;
   X[3022] := 3.2239845;
   X[3023] := 3.3288887;
   X[3024] := 3.4290748;
   X[3025] := 3.5245376;
   X[3026] := 3.6306174;
   X[3027] := 3.7275321;
   X[3028] := 3.8287132;
   X[3029] := 3.927261;
   X[3030] := 4.0291758;
   X[3031] := 4.1305375;
   X[3032] := 4.2238994;
   X[3033] := 4.3312664;
   X[3034] := 4.4264417;
   X[3035] := 4.526713;
   X[3036] := 4.6318994;
   X[3037] := 4.724176;
   X[3038] := 4.8276386;
   X[3039] := 4.928272;
   X[3040] := 5.0231757;
   X[3041] := 5.1239953;
   X[3042] := 5.223724;
   X[3043] := 5.323995;
   X[3044] := 5.424453;
   X[3045] := 5.525362;
   X[3046] := 5.6235485;
   X[3047] := 5.7188196;
   X[3048] := 5.8196335;
   X[3049] := 5.926277;
   X[3050] := 6.01749;
   X[3051] := 6.1050224;
   X[3052] := 6.1911025;
   X[3053] := 6.2721086;
   X[3054] := 6.350471;
   X[3055] := 6.4473224;
   X[3056] := 6.5459604;
   X[3057] := 6.6483274;
   X[3058] := 6.7456093;
   X[3059] := 6.8444285;
   X[3060] := 6.9463434;
   X[3061] := 7.0396147;
   X[3062] := 7.14262;
   X[3063] := 7.2407055;
   X[3064] := 7.3428917;
   X[3065] := 7.438078;
   X[3066] := 7.544721;
   X[3067] := 7.6421733;
   X[3068] := 7.736179;
   X[3069] := 7.8428063;
   X[3070] := 7.940365;
   X[3071] := 8.044456;
   X[3072] := 8.135737;
   X[3073] := 8.238105;
   X[3074] := 8.34528;
   X[3075] := 8.4401045;
   X[3076] := 8.535737;
   X[3077] := 8.635019;
   X[3078] := 8.740381;
   X[3079] := 8.841929;
   X[3080] := 8.935025;
   X[3081] := 9.034754;
   X[3082] := 9.136668;
   X[3083] := 9.237302;
   X[3084] := 9.332578;
   X[3085] := 9.434307;
   X[3086] := 9.53195;
   X[3087] := 9.640855;
   X[3088] := 9.736493;
   X[3089] := 9.832408;
   X[3090] := 9.930227;
   X[3091] := 10.039142;
   X[3092] := 10.131232;
   X[3093] := 10.231051;
   X[3094] := 10.330429;
   X[3095] := 10.432243;
   X[3096] := 10.529791;
   X[3097] := 10.63352;
   X[3098] := 10.733876;
   X[3099] := 10.828158;
   X[3100] := 10.927254;
   X[3101] := 11.023445;
   X[3102] := 11.128621;
   X[3103] := 11.228897;
   X[3104] := 11.324446;
   X[3105] := 11.423089;
   X[3106] := 11.521903;
   X[3107] := 11.629541;
   X[3108] := 11.722456;
   X[3109] := 11.822546;
   X[3110] := 11.922919;
   X[3111] := 12.019738;
   X[3112] := 12.121285;
   X[3113] := 12.221015;
   X[3114] := 12.31711;
   X[3115] := 12.422573;
   X[3116] := 12.522929;
   X[3117] := 12.618567;
   X[3118] := 12.724754;
   X[3119] := 12.81894;
   X[3120] := 12.915212;
   X[3121] := 13.016307;
   X[3122] := 13.118669;
   X[3123] := 13.216222;
   X[3124] := 13.316589;
   X[3125] := 13.4159565;
   X[3126] := 13.515318;
   X[3127] := 13.616505;
   X[3128] := 13.713776;
   X[3129] := 13.812414;
   X[3130] := 13.918695;
   X[3131] := 14.010786;
   X[3132] := 14.115153;
   X[3133] := 14.212973;
   X[3134] := 14.31043;
   X[3135] := 14.411978;
   X[3136] := 14.509345;
   X[3137] := 14.609526;
   X[3138] := 14.71144;
   X[3139] := 14.808989;
   X[3140] := 14.913802;
   X[3141] := 15.003371;
   X[3142] := 15.105467;
   X[3143] := 15.200116;
   X[3144] := 15.30068;
   X[3145] := 15.393058;
   X[3146] := 15.495165;
   X[3147] := 15.591356;
   X[3148] := 15.688271;
   X[3149] := 15.788569;
   X[3150] := 15.884032;
   X[3151] := 15.984958;
   X[3152] := 16.078962;
   X[3153] := 16.182436;
   X[3154] := 16.27391;
   X[3155] := 16.371006;
   X[3156] := 16.464664;
   X[3157] := 16.565943;
   X[3158] := 16.668139;
   X[3159] := 16.761145;
   X[3160] := 16.85689;
   X[3161] := 16.952633;
   X[3162] := 17.05729;
   X[3163] := 17.152203;
   X[3164] := 17.247038;
   X[3165] := 17.349602;
   X[3166] := 17.444431;
   X[3167] := 17.5408;
   X[3168] := 17.639996;
   X[3169] := 17.735012;
   X[3170] := 17.839931;
   X[3171] := 17.930767;
   X[3172] := 18.02815;
   X[3173] := 18.12698;
   X[3174] := 18.220715;
   X[3175] := 18.320364;
   X[3176] := 18.421837;
   X[3177] := 18.516758;
   X[3178] := 18.616045;
   X[3179] := 18.714157;
   X[3180] := 18.814072;
   X[3181] := 18.907455;
   X[3182] := 19.00029;
   X[3183] := 19.098295;
   X[3184] := 19.200663;
   X[3185] := 19.297142;
   X[3186] := 19.39788;
   X[3187] := 19.493801;
   X[3188] := 19.586275;
   X[3189] := 19.679651;
   X[3190] := 19.78603;
   X[3191] := 19.881477;
   X[3192] := 20.000278;
   X[3193] := 20.127155;
   X[3194] := 20.245878;
   X[3195] := 20.368128;
   X[3196] := 20.487148;
   X[3197] := 20.583235;
   X[3198] := 20.680521;
   X[3199] := 20.781872;
   X[3200] := 20.877792;
   X[3201] := 20.979069;
   X[3202] := 21.07743;
   X[3203] := 21.175076;
   X[3204] := 21.282347;
   X[3205] := 21.371809;
   X[3206] := 21.475542;
   X[3207] := 21.57118;
   X[3208] := 21.67291;
   X[3209] := 21.771357;
   X[3210] := 21.87109;
   X[3211] := 21.97191;
   X[3212] := 22.070745;
   X[3213] := 22.170372;
   X[3214] := 22.269379;
   X[3215] := 22.376106;
   X[3216] := 22.464926;
   X[3217] := 22.569479;
   X[3218] := 22.672384;
   X[3219] := 22.772305;
   X[3220] := 22.868128;
   X[3221] := 22.968937;
   X[3222] := 23.07058;
   X[3223] := 23.16358;
   X[3224] := 23.269947;
   X[3225] := 23.36205;
   X[3226] := 23.46433;
   X[3227] := 23.56532;
   X[3228] := 23.66333;
   X[3229] := 23.759235;
   X[3230] := 23.867155;
   X[3231] := 23.965612;
   X[3232] := 24.05716;
   X[3233] := 24.155884;
   X[3234] := 24.263342;
   X[3235] := 24.362442;
   X[3236] := 24.460714;
   X[3237] := 24.558176;
   X[3238] := 24.659628;
   X[3239] := 24.759459;
   X[3240] := 24.852186;
   X[3241] := 24.95391;
   X[3242] := 25.053635;
   X[3243] := 25.158182;
   X[3244] := 25.257915;
   X[3245] := 25.351559;
   X[3246] := 25.454927;
   X[3247] := 25.548931;
   X[3248] := 25.651932;
   X[3249] := 25.753654;
   X[3250] := 25.850208;
   X[3251] := 25.953394;
   X[3252] := 26.056581;
   X[3253] := 26.147043;
   X[3254] := 26.247953;
   X[3255] := 26.350044;
   X[3256] := 26.44714;
   X[3257] := 26.549511;
   X[3258] := 26.648325;
   X[3259] := 26.74906;
   X[3260] := 26.848692;
   X[3261] := 26.940432;
   X[3262] := 27.045975;
   X[3263] := 27.1418;
   X[3264] := 27.238708;
   X[3265] := 27.341171;
   X[3266] := 27.44381;
   X[3267] := 27.545267;
   X[3268] := 27.636906;
   X[3269] := 27.744719;
   X[3270] := 27.841002;
   X[3271] := 27.944555;
   X[3272] := 28.041187;
   X[3273] := 28.13265;
   X[3274] := 28.232927;
   X[3275] := 28.33283;
   X[3276] := 28.433384;
   X[3277] := 28.533842;
   X[3278] := 28.63248;
   X[3279] := 28.734396;
   X[3280] := 28.839396;
   X[3281] := 28.928768;
   X[3282] := 29.03231;
   X[3283] := 29.13304;
   X[3284] := 29.229507;
   X[3285] := 29.332235;
   X[3286] := 29.426598;
   X[3287] := 29.531965;
   X[3288] := 29.580423;
   X[3289] := 29.612755;
   X[3290] := 29.64728;
   X[3291] := 29.691607;
   X[3292] := 29.729671;
   X[3293] := 29.764744;
   X[3294] := 29.805613;
   X[3295] := 29.843763;
   X[3296] := 29.878738;
   X[3297] := 29.876654;
   X[3298] := 29.886017;
   X[3299] := 29.881754;
   X[3300] := 29.850193;
   X[3301] := 29.813211;
   X[3302] := 29.771793;
   X[3303] := 29.740717;
   X[3304] := 29.69848;
   X[3305] := 29.662506;
   X[3306] := 29.62344;
   X[3307] := 29.586565;
   X[3308] := 29.546526;
   X[3309] := 29.454744;
   X[3310] := 29.360846;
   X[3311] := 29.253382;
   X[3312] := 29.158281;
   X[3313] := 29.059101;
   X[3314] := 28.961727;
   X[3315] := 28.858818;
   X[3316] := 28.759722;
   X[3317] := 28.655186;
   X[3318] := 28.560537;
   X[3319] := 28.461723;
   X[3320] := 28.36126;
   X[3321] := 28.261084;
   X[3322] := 28.168255;
   X[3323] := 28.060797;
   X[3324] := 27.96107;
   X[3325] := 27.859068;
   X[3326] := 27.758966;
   X[3327] := 27.657244;
   X[3328] := 27.569328;
   X[3329] := 27.464962;
   X[3330] := 27.360596;
   X[3331] := 27.27241;
   X[3332] := 27.17177;
   X[3333] := 27.07177;
   X[3334] := 26.971313;
   X[3335] := 26.873674;
   X[3336] := 26.775764;
   X[3337] := 26.669403;
   X[3338] := 26.563574;
   X[3339] := 26.469482;
   X[3340] := 26.368025;
   X[3341] := 26.266478;
   X[3342] := 26.169834;
   X[3343] := 26.078472;
   X[3344] := 25.971563;
   X[3345] := 25.875004;
   X[3346] := 25.772552;
   X[3347] := 25.670004;
   X[3348] := 25.572638;
   X[3349] := 25.471632;
   X[3350] := 25.374456;
   X[3351] := 25.276903;
   X[3352] := 25.177631;
   X[3353] := 25.081078;
   X[3354] := 24.978525;
   X[3355] := 24.88443;
   X[3356] := 24.77652;
   X[3357] := 24.683344;
   X[3358] := 24.582062;
   X[3359] := 24.485147;
   X[3360] := 24.38487;
   X[3361] := 24.279062;
   X[3362] := 24.177961;
   X[3363] := 24.079689;
   X[3364] := 23.979599;
   X[3365] := 23.886322;
   X[3366] := 23.777233;
   X[3367] := 23.687593;
   X[3368] := 23.581488;
   X[3369] := 23.48604;
   X[3370] := 23.384127;
   X[3371] := 23.288488;
   X[3372] := 23.184212;
   X[3373] := 23.086834;
   X[3374] := 22.985659;
   X[3375] := 22.886477;
   X[3376] := 22.790104;
   X[3377] := 22.686556;
   X[3378] := 22.58629;
   X[3379] := 22.488918;
   X[3380] := 22.3941;
   X[3381] := 22.29236;
   X[3382] := 22.189919;
   X[3383] := 22.092999;
   X[3384] := 21.994902;
   X[3385] := 21.893812;
   X[3386] := 21.792625;
   X[3387] := 21.694088;
   X[3388] := 21.59235;
   X[3389] := 21.49863;
   X[3390] := 21.397068;
   X[3391] := 21.293348;
   X[3392] := 21.196524;
   X[3393] := 21.0997;
   X[3394] := 20.9947;
   X[3395] := 20.89579;
   X[3396] := 20.798689;
   X[3397] := 20.701242;
   X[3398] := 20.600412;
   X[3399] := 20.503046;
   X[3400] := 20.401136;
   X[3401] := 20.294594;
   X[3402] := 20.20195;
   X[3403] := 20.105131;
   X[3404] := 20.002398;
   X[3405] := 19.90676;
   X[3406] := 19.800934;
   X[3407] := 19.703669;
   X[3408] := 19.60539;
   X[3409] := 19.506657;
   X[3410] := 19.404295;
   X[3411] := 19.305471;
   X[3412] := 19.206018;
   X[3413] := 19.112652;
   X[3414] := 19.010918;
   X[3415] := 18.905918;
   X[3416] := 18.809828;
   X[3417] := 18.712456;
   X[3418] := 18.610184;
   X[3419] := 18.504637;
   X[3420] := 18.40754;
   X[3421] := 18.311901;
   X[3422] := 18.207354;
   X[3423] := 18.116348;
   X[3424] := 18.010445;
   X[3425] := 17.914625;
   X[3426] := 17.8138;
   X[3427] := 17.713434;
   X[3428] := 17.611885;
   X[3429] := 17.511248;
   X[3430] := 17.422699;
   X[3431] := 17.313423;
   X[3432] := 17.213789;
   X[3433] := 17.11069;
   X[3434] := 17.015944;
   X[3435] := 16.91578;
   X[3436] := 16.816774;
   X[3437] := 16.716045;
   X[3438] := 16.621677;
   X[3439] := 16.515497;
   X[3440] := 16.415758;
   X[3441] := 16.315577;
   X[3442] := 16.212849;
   X[3443] := 16.128843;
   X[3444] := 16.02339;
   X[3445] := 15.920018;
   X[3446] := 15.821662;
   X[3447] := 15.727843;
   X[3448] := 15.625742;
   X[3449] := 15.526646;
   X[3450] := 15.431284;
   X[3451] := 15.33055;
   X[3452] := 15.230816;
   X[3453] := 15.1187315;
   X[3454] := 15.024918;
   X[3455] := 14.924635;
   X[3456] := 14.825279;
   X[3457] := 14.73154;
   X[3458] := 14.630268;
   X[3459] := 14.527444;
   X[3460] := 14.42462;
   X[3461] := 14.332257;
   X[3462] := 14.229896;
   X[3463] := 14.1328;
   X[3464] := 14.029524;
   X[3465] := 13.936518;
   X[3466] := 13.832422;
   X[3467] := 13.732518;
   X[3468] := 13.632332;
